{region 'Documentation'}
(*!
<summary>Checks exact finding count and identities; at most one finding per subject.</summary>
*)
{endregion}
METHOD PRIVATE CheckFindings
VAR
    Index : UINT;
    Matches : BOOL;
END_VAR
Index := 1;
FFindingsMatch := TRUE;
Matches := CheckFinding(Subject := FEqual,
    ExpectedResult := FEqualExpectedResult,
    ExpectedFinding := FEqualExpectedFinding,
    Index := Index);
FFindingsMatch := FFindingsMatch AND Matches;
Matches := CheckFinding(Subject := FPattern,
    ExpectedResult := FPatternExpectedResult,
    ExpectedFinding := FPatternExpectedFinding,
    Index := Index);
FFindingsMatch := FFindingsMatch AND Matches;
Matches := CheckFinding(Subject := FAll,
    ExpectedResult := FAllExpectedResult,
    ExpectedFinding := FAllExpectedFinding,
    Index := Index);
FFindingsMatch := FFindingsMatch AND Matches;
Matches := CheckFinding(Subject := FValue,
    ExpectedResult := FValueExpectedResult,
    ExpectedFinding := FValueExpectedFinding,
    Index := Index);
FFindingsMatch := FFindingsMatch AND Matches;
FFindingsMatch := FFindingsMatch
    AND (FCaptureStatus.SequenceId = UINT_TO_UDINT(Index - 1))
    AND (FCaptureStatus.LostEventCount = 0);
END_METHOD

{region 'Documentation'}
(*!
<summary>Rejects incomplete subject, capture or outer Assertion setup.</summary>
*)
{endregion}
METHOD PROTECTED CheckInitialization : BOOL //! TRUE when the inherited initialization check and this concrete fixture check both accept the setup.
CheckInitialization := SUPER^.CheckInitialization();
IF NOT CheckInitialization THEN
    RETURN;
END_IF;

CheckInitialization := FSetupValid
    AND FResults.IsInitialized
    AND FActivity.IsInitialized
    AND FInputs.IsInitialized
    AND FFindings.IsInitialized;
IF NOT CheckInitialization THEN
    EventPublisher.PublishEvent(Event := CreateFrameworkEvent(Name := Name,
        ResourceName := '',
        State := State,
        Severity := E_EventSeverity.Error,
        Message := 'Array selftest setup failed.'));
END_IF;
END_METHOD

{region 'Documentation'}
(*!
<summary>Verifies input preservation without using the tested comparison algorithm.</summary>
*)
{endregion}
METHOD PRIVATE CheckInputs
VAR
    Index : DINT;
    ActualBits : FloatingPointBits_Real;
    SavedBits : FloatingPointBits_Real;
    WideActualBits : FloatingPointBits_LReal;
    WideSavedBits : FloatingPointBits_LReal;
END_VAR
FInputsMatch := TRUE;
FOR Index := -2 TO 1 DO
    ActualBits.Value := FData[Index];
    SavedBits.Value := FDataBefore[Index];
    WideActualBits.Value := FWideData[Index];
    WideSavedBits.Value := FWideDataBefore[Index];
    FInputsMatch := FInputsMatch
        AND (ActualBits.Bits = SavedBits.Bits)
        AND (WideActualBits.Bits = WideSavedBits.Bits);
END_FOR;
FOR Index := 4 TO 5 DO
    ActualBits.Value := FExpected[Index];
    SavedBits.Value := FExpectedBefore[Index];
    FInputsMatch := FInputsMatch AND (ActualBits.Bits = SavedBits.Bits);
END_FOR;
END_METHOD

{region 'Documentation'}
(*!
<summary>Checks literal evaluation results, or NotEvaluated on the reset call.</summary>
*)
{endregion}
METHOD PRIVATE CheckResults
IF FEvaluateSubjects THEN
    FResultsMatch := (FEqual.Result = FEqualExpectedResult)
        AND (FPattern.Result = FPatternExpectedResult)
        AND (FAll.Result = FAllExpectedResult)
        AND (FValue.Result = FValueExpectedResult);
ELSE
    FResultsMatch := (FEqual.Result = E_Result.NotEvaluated)
        AND (FPattern.Result = E_Result.NotEvaluated)
        AND (FAll.Result = E_Result.NotEvaluated)
        AND (FValue.Result = E_Result.NotEvaluated);
END_IF;
FActivityMatch := (FEqual.Enabled = FSubjectEnable)
    AND (FEqual.ObservationActive = (FEvaluateSubjects AND FSubjectEnable))
    AND (FEqual.EvaluationActive = (FEvaluateSubjects AND FSubjectEnable))
    AND (FPattern.Enabled = FSubjectEnable)
    AND (FPattern.ObservationActive = (FEvaluateSubjects AND FSubjectEnable))
    AND (FPattern.EvaluationActive = (FEvaluateSubjects AND FSubjectEnable))
    AND (FAll.Enabled = FSubjectEnable)
    AND (FAll.ObservationActive = (FEvaluateSubjects AND FSubjectEnable))
    AND (FAll.EvaluationActive = (FEvaluateSubjects AND FSubjectEnable))
    AND (FValue.Enabled = FSubjectEnable)
    AND (FValue.ObservationActive = (FEvaluateSubjects AND FSubjectEnable))
    AND (FValue.EvaluationActive = (FEvaluateSubjects AND FSubjectEnable));
END_METHOD

{region 'Documentation'}
(*!
<summary>Initializes outer checks and isolates intentional subject findings.</summary>
*)
{endregion}
METHOD PROTECTED Configure
VAR
    Initialized : BOOL;
END_VAR
FPreparationStateCount := 0;
FTestStateCount := 1;
FResults.Initialize(Parent := THIS^,
    AssertionName := 'Results');
FActivity.Initialize(Parent := THIS^,
    AssertionName := 'Activity');
FInputs.Initialize(Parent := THIS^,
    AssertionName := 'Inputs');
FFindings.Initialize(Parent := THIS^,
    AssertionName := 'Findings');
FSetupValid := FCapture.Initialize(Buffer := FEvents,
    FifoControl := FCaptureFifo,
    Status := FCaptureStatus);
FEqual.BindPublisher(Publisher := FCapture);
Initialized := FEqual.Initialize(Parent := THIS^,
    AssertionName := 'Equal');
FSetupValid := FSetupValid AND Initialized;
FPattern.BindPublisher(Publisher := FCapture);
Initialized := FPattern.Initialize(Parent := THIS^,
    AssertionName := 'Pattern');
FSetupValid := FSetupValid AND Initialized;
FAll.BindPublisher(Publisher := FCapture);
Initialized := FAll.Initialize(Parent := THIS^,
    AssertionName := 'All');
FSetupValid := FSetupValid AND Initialized;
FValue.BindPublisher(Publisher := FCapture);
Initialized := FValue.Initialize(Parent := THIS^,
    AssertionName := 'Value');
FSetupValid := FSetupValid AND Initialized;
END_METHOD

{region 'Documentation'}
(*!
<summary>Completes abort; no asynchronous resource is owned.</summary>
*)
{endregion}
METHOD PROTECTED ProcessAbort
VAR_INPUT
    Enable : BOOL; //! Phase permission supplied by the owning Test Case; FALSE does not authorize progression, while observation may continue.
END_VAR
IF Enable THEN
    CompleteAbort();
END_IF;
END_METHOD

{region 'Documentation'}
(*!
<summary>Latches this call's checks before progression is permitted.</summary>
*)
{endregion}
METHOD PROTECTED ProcessAssertions
VAR_INPUT
    Enable : BOOL; //! Phase permission supplied by the owning Test Case; FALSE does not authorize progression, while observation may continue.
END_VAR
VAR
    Check : BOOL;
END_VAR
Check := Enable AND FObservationReady;
FResults(Enable := Check,
    State := State,
    IN := FResultsMatch);
FActivity(Enable := Check,
    State := State,
    IN := FActivityMatch);
FInputs(Enable := Check,
    State := State,
    IN := FInputsMatch);
FFindings(Enable := Check,
    State := State,
    IN := FFindingsMatch);
IF Check THEN
    FChecked := TRUE;
END_IF;
END_METHOD

{region 'Documentation'}
(*!
<summary>No Preparation phase is needed.</summary>
*)
{endregion}
METHOD PROTECTED ProcessPreparations
VAR_INPUT
    // SA0033: Required hook; this test has no Preparation phase.
    {attribute 'analysis' := '-33'}
    Enable : BOOL; //! Phase permission supplied by the owning Test Case; FALSE does not authorize progression, while observation may continue.
END_VAR
END_METHOD

{region 'Documentation'}
(*!
<summary>Restarts the scenario sequence and outer checks.</summary>
*)
{endregion}
METHOD PROTECTED ProcessReset
FScenario := ScenarioFiniteEqual;
FChecked := FALSE;
FSubjectEnable := FALSE;
FEvaluateSubjects := FALSE;
FObservationReady := FALSE;
FFirstFailedScenario := 0;
FFailedDuringEvaluation := FALSE;
FCapture.Reset();
ResetSubjects();
FResults.Reset();
FActivity.Reset();
FInputs.Reset();
FFindings.Reset();
CompleteReset();
END_METHOD

{region 'Documentation'}
(*!
<summary>Consumes reset, evaluates, then waits for the outer checks before advancing.</summary>
*)
{endregion}
METHOD PROTECTED ProcessTests
VAR_INPUT
    Enable : BOOL; //! Phase permission supplied by the owning Test Case; FALSE does not authorize progression, while observation may continue.
END_VAR
IF NOT Enable THEN
    RETURN;
END_IF;

IF FChecked THEN
    FChecked := FALSE;
    FObservationReady := FALSE;
    IF FEvaluateSubjects THEN
        IF FScenario = LastScenario THEN
            CompleteTests();
            RETURN;
        END_IF;
        FScenario := FScenario + 1;
    END_IF;
    FEvaluateSubjects := NOT FEvaluateSubjects;
END_IF;

IF NOT SelectScenario() THEN
    RETURN;
END_IF;
FCapture.Reset();
IF NOT FEvaluateSubjects THEN
    ResetSubjects();
END_IF;
FDataBefore := FData;
FExpectedBefore := FExpected;
FWideDataBefore := FWideData;

CallSubjects();
CheckResults();
CheckInputs();
CheckFindings();
IF (FFirstFailedScenario = 0)
    AND NOT (FResultsMatch AND FActivityMatch AND FInputsMatch AND FFindingsMatch) THEN
    FFirstFailedScenario := FScenario;
    FFailedDuringEvaluation := FEvaluateSubjects;
END_IF;
FObservationReady := TRUE;
END_METHOD

{region 'Documentation'}
(*!
<summary>Queues reset; the next bound FB call consumes it without evaluating.</summary>
*)
{endregion}
METHOD PRIVATE ResetSubjects
FEqual.Reset();
FPattern.Reset();
FAll.Reset();
FValue.Reset();
END_METHOD

{region 'Documentation'}
(*!
<summary>Selects explicit stimuli and expected results for one scenario.</summary>
*)
{endregion}
METHOD PRIVATE SelectScenario : BOOL //! TRUE after selecting a supported scenario and its literal expectations; FALSE reports an unknown scenario.
VAR
    Index : DINT;
END_VAR
SelectScenario := FALSE;
FSubjectEnable := TRUE;
FQuietNaN.Bits := QuietNaNBits;
FPositiveInfinity.Bits := PositiveInfinityBits;
FNegativeInfinity.Bits := NegativeInfinityBits;
FWideQuietNaN.Bits := WideQuietNaNBits;
FWidePositiveInfinity.Bits := WidePositiveInfinityBits;
FWideNegativeInfinity.Bits := WideNegativeInfinityBits;
FActual := 1.0;
FReference := 1.0;
FWideActual := 1.0;
FWideExpected := 1.0;
FTolerance := 0.0;
FWideTolerance := 0.0;
CASE FScenario OF
    ScenarioFiniteEqual:
        FEqualExpectedResult := E_Result.Passed;
        FEqualExpectedFinding := FALSE;
        FPatternExpectedResult := E_Result.Passed;
        FPatternExpectedFinding := FALSE;
        FAllExpectedResult := E_Result.Passed;
        FAllExpectedFinding := FALSE;
        FValueExpectedResult := E_Result.Passed;
        FValueExpectedFinding := FALSE;
    ScenarioToleranceBoundary:
        FActual := 1.25;
        FWideActual := 1.25;
        FTolerance := 0.25;
        FWideTolerance := 0.25;
        FEqualExpectedResult := E_Result.Passed;
        FEqualExpectedFinding := FALSE;
        FPatternExpectedResult := E_Result.Passed;
        FPatternExpectedFinding := FALSE;
        FAllExpectedResult := E_Result.Passed;
        FAllExpectedFinding := FALSE;
        FValueExpectedResult := E_Result.Passed;
        FValueExpectedFinding := FALSE;
    ScenarioOutsideTolerance:
        FActual := 1.5;
        FWideActual := 1.5;
        FTolerance := 0.25;
        FWideTolerance := 0.25;
        FEqualExpectedResult := E_Result.Failed;
        FEqualExpectedFinding := TRUE;
        FPatternExpectedResult := E_Result.Failed;
        FPatternExpectedFinding := TRUE;
        FAllExpectedResult := E_Result.Failed;
        FAllExpectedFinding := TRUE;
        FValueExpectedResult := E_Result.Failed;
        FValueExpectedFinding := TRUE;
    ScenarioNaNBeforeValidMatch:
        FEqualExpectedResult := E_Result.Failed;
        FEqualExpectedFinding := TRUE;
        FPatternExpectedResult := E_Result.Passed;
        FPatternExpectedFinding := FALSE;
        FAllExpectedResult := E_Result.Failed;
        FAllExpectedFinding := TRUE;
        FValueExpectedResult := E_Result.Passed;
        FValueExpectedFinding := FALSE;
    ScenarioOnlyNaNActual:
        FActual := FQuietNaN.Value;
        FWideActual := FWideQuietNaN.Value;
        FEqualExpectedResult := E_Result.Failed;
        FEqualExpectedFinding := TRUE;
        FPatternExpectedResult := E_Result.Failed;
        FPatternExpectedFinding := TRUE;
        FAllExpectedResult := E_Result.Failed;
        FAllExpectedFinding := TRUE;
        FValueExpectedResult := E_Result.Failed;
        FValueExpectedFinding := TRUE;
    ScenarioPositiveInfinityMatch:
        FActual := FPositiveInfinity.Value;
        FReference := FPositiveInfinity.Value;
        FWideActual := FWidePositiveInfinity.Value;
        FWideExpected := FWidePositiveInfinity.Value;
        FEqualExpectedResult := E_Result.Error;
        FEqualExpectedFinding := TRUE;
        FPatternExpectedResult := E_Result.Passed;
        FPatternExpectedFinding := FALSE;
        FAllExpectedResult := E_Result.Passed;
        FAllExpectedFinding := FALSE;
        FValueExpectedResult := E_Result.Passed;
        FValueExpectedFinding := FALSE;
    ScenarioNegativeInfinityMatch:
        FActual := FNegativeInfinity.Value;
        FReference := FNegativeInfinity.Value;
        FWideActual := FWideNegativeInfinity.Value;
        FWideExpected := FWideNegativeInfinity.Value;
        FEqualExpectedResult := E_Result.Error;
        FEqualExpectedFinding := TRUE;
        FPatternExpectedResult := E_Result.Passed;
        FPatternExpectedFinding := FALSE;
        FAllExpectedResult := E_Result.Passed;
        FAllExpectedFinding := FALSE;
        FValueExpectedResult := E_Result.Passed;
        FValueExpectedFinding := FALSE;
    ScenarioOppositeInfinities:
        FActual := FPositiveInfinity.Value;
        FReference := FNegativeInfinity.Value;
        FWideActual := FWidePositiveInfinity.Value;
        FWideExpected := FWideNegativeInfinity.Value;
        FEqualExpectedResult := E_Result.Error;
        FEqualExpectedFinding := TRUE;
        FPatternExpectedResult := E_Result.Failed;
        FPatternExpectedFinding := TRUE;
        FAllExpectedResult := E_Result.Failed;
        FAllExpectedFinding := TRUE;
        FValueExpectedResult := E_Result.Failed;
        FValueExpectedFinding := TRUE;
    ScenarioPositiveInfinityActual:
        FActual := FPositiveInfinity.Value;
        FWideActual := FWidePositiveInfinity.Value;
        FEqualExpectedResult := E_Result.Failed;
        FEqualExpectedFinding := TRUE;
        FPatternExpectedResult := E_Result.Failed;
        FPatternExpectedFinding := TRUE;
        FAllExpectedResult := E_Result.Failed;
        FAllExpectedFinding := TRUE;
        FValueExpectedResult := E_Result.Failed;
        FValueExpectedFinding := TRUE;
    ScenarioNegativeInfinityActual:
        FActual := FNegativeInfinity.Value;
        FWideActual := FWideNegativeInfinity.Value;
        FEqualExpectedResult := E_Result.Failed;
        FEqualExpectedFinding := TRUE;
        FPatternExpectedResult := E_Result.Failed;
        FPatternExpectedFinding := TRUE;
        FAllExpectedResult := E_Result.Failed;
        FAllExpectedFinding := TRUE;
        FValueExpectedResult := E_Result.Failed;
        FValueExpectedFinding := TRUE;
    ScenarioNaNExpected:
        FReference := FQuietNaN.Value;
        FWideExpected := FWideQuietNaN.Value;
        FEqualExpectedResult := E_Result.Error;
        FEqualExpectedFinding := TRUE;
        FPatternExpectedResult := E_Result.Error;
        FPatternExpectedFinding := TRUE;
        FAllExpectedResult := E_Result.Error;
        FAllExpectedFinding := TRUE;
        FValueExpectedResult := E_Result.Error;
        FValueExpectedFinding := TRUE;
    ScenarioLateNaNExpected:
        FEqualExpectedResult := E_Result.Error;
        FEqualExpectedFinding := TRUE;
        FPatternExpectedResult := E_Result.Error;
        FPatternExpectedFinding := TRUE;
        FAllExpectedResult := E_Result.Passed;
        FAllExpectedFinding := FALSE;
        FValueExpectedResult := E_Result.Passed;
        FValueExpectedFinding := FALSE;
    ScenarioNegativeTolerance:
        FTolerance := -0.25;
        FWideTolerance := -0.25;
        FEqualExpectedResult := E_Result.Error;
        FEqualExpectedFinding := TRUE;
        FPatternExpectedResult := E_Result.Error;
        FPatternExpectedFinding := TRUE;
        FAllExpectedResult := E_Result.Error;
        FAllExpectedFinding := TRUE;
        FValueExpectedResult := E_Result.Error;
        FValueExpectedFinding := TRUE;
    ScenarioNaNTolerance:
        FTolerance := FQuietNaN.Value;
        FWideTolerance := FWideQuietNaN.Value;
        FEqualExpectedResult := E_Result.Error;
        FEqualExpectedFinding := TRUE;
        FPatternExpectedResult := E_Result.Error;
        FPatternExpectedFinding := TRUE;
        FAllExpectedResult := E_Result.Error;
        FAllExpectedFinding := TRUE;
        FValueExpectedResult := E_Result.Error;
        FValueExpectedFinding := TRUE;
    ScenarioInfiniteTolerance:
        FTolerance := FPositiveInfinity.Value;
        FWideTolerance := FWidePositiveInfinity.Value;
        FEqualExpectedResult := E_Result.Error;
        FEqualExpectedFinding := TRUE;
        FPatternExpectedResult := E_Result.Error;
        FPatternExpectedFinding := TRUE;
        FAllExpectedResult := E_Result.Error;
        FAllExpectedFinding := TRUE;
        FValueExpectedResult := E_Result.Error;
        FValueExpectedFinding := TRUE;
ELSE
    Error(Message := 'Unknown array Assertion scenario.');
    RETURN;
END_CASE;
FOR Index := -2 TO 1 DO
    FData[Index] := FActual;
    FWideData[Index] := FWideActual;
END_FOR;
FExpected[4] := FReference;
FExpected[5] := FReference;
IF FScenario = ScenarioNaNBeforeValidMatch THEN
    FData[-2] := FQuietNaN.Value;
    FWideData[-2] := FWideQuietNaN.Value;
END_IF;
IF FScenario = ScenarioLateNaNExpected THEN
    FExpected[5] := FQuietNaN.Value;
    FData[-2] := 9.0;
END_IF;
SelectScenario := TRUE;
END_METHOD

END_FUNCTION_BLOCK

// ---- Framework/Assertions/POU/Arrays/Real/AssertEqualArray_Real.TcPOU
{region 'Documentation'}
(*!
<summary>Compares the entire Expected array with IN starting at StartIndex.</summary>
<description>

StartIndex is an absolute declared IN index. The entire Expected array, starting at its
own lower bound, determines the compared length and must fit IN. Invalid references or ranges
report Error.

Keep supplied arrays stable for the call. Input data is read, not copied or retained as a
snapshot.

Every Expected element must be finite; otherwise Error. A non-finite actual element is a
mismatch (Failed), not an invalid Expected value.

Tolerance is absolute, in the same units as the values, finite and non-negative. Its
default zero requests exact comparison. The equality boundary is inclusive; larger differences
are unequal. Difference checking avoids overflow for large finite operands.

Numeric diagnostics use the formatter's default six significant digits; rounding affects
the message only, not the comparison.

</description>
*)
{endregion}
FUNCTION_BLOCK AssertEqualArray_Real EXTENDS AssertionBase
VAR_INPUT
    Tolerance : REAL := 0.0; //! Maximum absolute allowed difference; finite and non-negative.
    StartIndex : DINT; //! First compared index in IN; Expected starts at its own lower bound.
END_VAR
VAR_IN_OUT CONSTANT
    IN : ARRAY[*] OF REAL; //! Read-only actual data; the selected range must remain stable during the call.
    Expected : ARRAY[*] OF REAL; //! Read-only expected sequence starting at its own lower bound; must fit the selected actual range.
END_VAR

SUPER^();

{region 'Documentation'}
(*!
<summary>Validate the selected range and expectations before comparing elements.</summary>
*)
{endregion}
METHOD PROTECTED Assert
VAR
    ReferenceValue : REAL;
    ValuesEqual : BOOL;
    Value : REAL;
    InLowerIndex : DINT;
    InUpperIndex : DINT;
    ExpectedLowerIndex : DINT;
    ExpectedUpperIndex : DINT;
    ExpectedLength : LINT;
    EndIndex : LINT;
    Offset : LINT;
    InIndex : DINT;
    ExpectedIndex : DINT;
    Message : STRING(GVL_Constants.MessageLength);
    ExpectedText : STRING(GVL_Constants.AssertionValueLength);
    ActualText : STRING(GVL_Constants.AssertionValueLength);
END_VAR
IF NOT EvaluationActive THEN
    RETURN;
END_IF;

IF Result = E_Result.Error THEN
    RETURN;
END_IF;

// C0371: FB inputs are checked here before any reference access.
{warning disable C0371}
IF NOT __ISVALIDREF(IN) THEN
    Error(Message := 'Assertion error: IN reference is invalid.');
    RETURN;
END_IF;

IF NOT __ISVALIDREF(Expected) THEN
    Error(Message := 'Assertion error: Expected reference is invalid.');
    RETURN;
END_IF;

IF NOT Tc2_Utilities.RealIsFinite(x := Tolerance) THEN
    Error(Message := 'Assertion error: Tolerance must be finite.');
    RETURN;
END_IF;

IF Tolerance < 0.0 THEN
    Error(Message := 'Assertion error: Tolerance must not be negative.');
    RETURN;
END_IF;

InLowerIndex := LOWER_BOUND(IN, 1);
InUpperIndex := UPPER_BOUND(IN, 1);
ExpectedLowerIndex := LOWER_BOUND(Expected, 1);
ExpectedUpperIndex := UPPER_BOUND(Expected, 1);
ExpectedLength := DINT_TO_LINT(ExpectedUpperIndex) - DINT_TO_LINT(ExpectedLowerIndex) + 1;
EndIndex := DINT_TO_LINT(StartIndex) + ExpectedLength - 1;

IF (ExpectedLength <= 0)
    OR (StartIndex < InLowerIndex) OR (StartIndex > InUpperIndex)
    OR (EndIndex > DINT_TO_LINT(InUpperIndex)) THEN
    Message := CONCAT('Assertion error: array range is invalid. StartIndex = ',
        DINT_TO_STRING(StartIndex));
    Message := CONCAT(Message, ', EndIndex = ');
    Message := CONCAT(Message, LINT_TO_STRING(EndIndex));
    Message := CONCAT(Message, ', InLowerIndex = ');
    Message := CONCAT(Message, DINT_TO_STRING(InLowerIndex));
    Message := CONCAT(Message, ', InUpperIndex = ');
    Message := CONCAT(Message, DINT_TO_STRING(InUpperIndex));
    Message := CONCAT(Message, ', ExpectedLength = ');
    Message := CONCAT(Message, LINT_TO_STRING(ExpectedLength));
    Message := CONCAT(Message, '.');
    Error(Message := Message);
    RETURN;
END_IF;

FOR Offset := 0 TO ExpectedLength - 1 DO
    ExpectedIndex := LINT_TO_DINT(DINT_TO_LINT(ExpectedLowerIndex) + Offset);
    Value := Expected[ExpectedIndex];
    IF NOT Tc2_Utilities.RealIsFinite(x := Value) THEN
        Message := CONCAT('Assertion error: Expected element must be finite. Index = ',
            DINT_TO_STRING(ExpectedIndex));
        Message := CONCAT(Message, '.');
        Error(Message := Message);
        RETURN;
    END_IF;
END_FOR;

IF Result = E_Result.Failed THEN
    RETURN;
END_IF;

FOR Offset := 0 TO ExpectedLength - 1 DO
    InIndex := LINT_TO_DINT(DINT_TO_LINT(StartIndex) + Offset);
    ExpectedIndex := LINT_TO_DINT(DINT_TO_LINT(ExpectedLowerIndex) + Offset);
    Value := IN[InIndex];
    ReferenceValue := Expected[ExpectedIndex];
    ValuesEqual := FALSE;
    IF NOT Tc2_Utilities.RealIsNaN(x := Value) THEN
        IF Value = ReferenceValue THEN
            ValuesEqual := TRUE;
        ELSIF Tc2_Utilities.RealIsFinite(x := Value)
            AND Tc2_Utilities.RealIsFinite(x := ReferenceValue) THEN
            ValuesEqual := IsWithinTolerance_Real(IN := Value,
                Expected := ReferenceValue,
                Tolerance := Tolerance);
        END_IF;
    END_IF;
    IF NOT ValuesEqual THEN
        ExpectedText := CreateAssertionTextValue_Real(Value := Expected[ExpectedIndex]);
        Value := IN[InIndex];
        IF Tc2_Utilities.RealIsFinite(x := Value) THEN
            ActualText := CreateAssertionTextValue_Real(Value := IN[InIndex]);
        ELSE
            ActualText := '<non-finite>';
        END_IF;
        Message := CONCAT('Assertion failed: array elements differ. Expected[',
            DINT_TO_STRING(ExpectedIndex));
        Message := CONCAT(Message, '] = ');
        Message := CONCAT(Message, ExpectedText);
        Message := CONCAT(Message, ', IN[');
        Message := CONCAT(Message, DINT_TO_STRING(InIndex));
        Message := CONCAT(Message, '] = ');
        Message := CONCAT(Message, ActualText);
        Message := CONCAT(Message, '.');
        Message := CONCAT(Message, ' Tolerance = ');
        Message := CONCAT(Message, CreateAssertionTextValue_Real(Value := Tolerance));
        Fail(Message := Message);
        RETURN;
    END_IF;
END_FOR;

Pass();
{warning restore C0371}
END_METHOD

END_FUNCTION_BLOCK

// ---- Framework/Assertions/POU/Arrays/Real/AssertArrayContainsArray_Real.TcPOU
{region 'Documentation'}
(*!
<summary>Searches the selected IN range for the complete contiguous Expected pattern.</summary>
<description>

StartIndex is an absolute declared IN index, not an offset. Length selects 1..255
elements; the complete selected range must fit IN. Invalid references or ranges report
Error.

Keep supplied arrays stable for the call. Input data is read, not copied or retained as a
snapshot.

The complete Expected pattern must be nonempty and fit the selected IN range; an
oversized pattern reports Error, not a missing-match result.

Expected must not contain NaN (Error), but may contain either infinity. Actual NaN never
matches; equal signed infinities match. Non-finite data elsewhere in a search does not
invalidate the entire range.

Tolerance is absolute, in the same units as the values, finite and non-negative. Its
default zero requests exact comparison. The equality boundary is inclusive; larger differences
are unequal. Difference checking avoids overflow for large finite operands.

Numeric diagnostics use the formatter's default six significant digits; rounding affects
the message only, not the comparison.

</description>
*)
{endregion}
FUNCTION_BLOCK AssertArrayContainsArray_Real EXTENDS AssertionBase
VAR_INPUT
    StartIndex : DINT; //! First selected index in IN; uses the array's declared index range, not a zero-based offset.
    Length : USINT; //! Number of searched elements, from 1 through 255.
    Tolerance : REAL := 0.0; //! Maximum absolute difference accepted as equal; must be finite and non-negative.
END_VAR
VAR_IN_OUT CONSTANT
    IN : ARRAY[*] OF REAL; //! Read-only search data; keep stable during the call.
    Expected : ARRAY[*] OF REAL; //! Read-only expected sequence starting at its own lower bound; must fit the selected actual range.
END_VAR

SUPER^();

{region 'Documentation'}
(*!
<summary>Validate configuration before searching the selected range.</summary>
*)
{endregion}
METHOD PROTECTED Assert
VAR
    InLowerIndex : DINT;
    InUpperIndex : DINT;
    EndIndex : LINT;
    Offset : LINT;
    InIndex : DINT;
    ExpectedLowerIndex : DINT;
    ExpectedUpperIndex : DINT;
    ExpectedLength : LINT;
    ExpectedIndex : DINT;
    CandidateOffset : LINT;
    PatternFound : BOOL;
    PatternMatches : BOOL;
    ValuesEqual : BOOL;
    ExpectedValue : REAL;
    Message : STRING(GVL_Constants.MessageLength);
    Value : REAL;
END_VAR
IF NOT EvaluationActive THEN
    RETURN;
END_IF;

IF Result = E_Result.Error THEN
    RETURN;
END_IF;

// C0371: FB input is checked here before any reference access.
{warning disable C0371}
IF NOT __ISVALIDREF(IN) THEN
    Error(Message := 'Assertion error: IN reference is invalid.');
    RETURN;
END_IF;

IF NOT Tc2_Utilities.RealIsFinite(x := Tolerance) THEN
    Error(Message := 'Assertion error: Tolerance must be finite.');
    RETURN;
END_IF;

IF Tolerance < 0.0 THEN
    Error(Message := 'Assertion error: Tolerance must not be negative.');
    RETURN;
END_IF;

IF NOT __ISVALIDREF(Expected) THEN
    Error(Message := 'Assertion error: Expected reference is invalid.');
    RETURN;
END_IF;

InLowerIndex := LOWER_BOUND(IN, 1);
InUpperIndex := UPPER_BOUND(IN, 1);
EndIndex := DINT_TO_LINT(StartIndex) + USINT_TO_LINT(Length) - 1;

ExpectedLowerIndex := LOWER_BOUND(Expected, 1);
ExpectedUpperIndex := UPPER_BOUND(Expected, 1);
ExpectedLength := DINT_TO_LINT(ExpectedUpperIndex) - DINT_TO_LINT(ExpectedLowerIndex) + 1;

IF (Length = 0)
    OR (ExpectedLength <= 0) OR (ExpectedLength > USINT_TO_LINT(Length))
    OR (StartIndex < InLowerIndex) OR (StartIndex > InUpperIndex)
    OR (EndIndex > DINT_TO_LINT(InUpperIndex)) THEN
    Message := CONCAT('Assertion error: array range or pattern is invalid. StartIndex = ',
        DINT_TO_STRING(StartIndex));
    Message := CONCAT(Message, ', Length = ');
    Message := CONCAT(Message, USINT_TO_STRING(Length));
    Message := CONCAT(Message, ', ExpectedLength = ');
    Message := CONCAT(Message, LINT_TO_STRING(ExpectedLength));
    Message := CONCAT(Message, '.');
    Error(Message := Message);
    RETURN;
END_IF;

FOR Offset := 0 TO ExpectedLength - 1 DO
    ExpectedIndex := LINT_TO_DINT(DINT_TO_LINT(ExpectedLowerIndex) + Offset);
    ExpectedValue := Expected[ExpectedIndex];
    IF Tc2_Utilities.RealIsNaN(x := ExpectedValue) THEN
        Message := CONCAT('Assertion error: Expected must not contain NaN. Index = ',
            DINT_TO_STRING(ExpectedIndex));
        Error(Message := Message);
        RETURN;
    END_IF;
END_FOR;

IF Result = E_Result.Failed THEN
    RETURN;
END_IF;

PatternFound := FALSE;
FOR CandidateOffset := 0 TO USINT_TO_LINT(Length) - ExpectedLength DO
    PatternMatches := TRUE;
    FOR Offset := 0 TO ExpectedLength - 1 DO
        InIndex := LINT_TO_DINT(DINT_TO_LINT(StartIndex) + CandidateOffset + Offset);
        ExpectedIndex := LINT_TO_DINT(DINT_TO_LINT(ExpectedLowerIndex) + Offset);
        Value := IN[InIndex];
        ExpectedValue := Expected[ExpectedIndex];
        ValuesEqual := FALSE;
        IF NOT Tc2_Utilities.RealIsNaN(x := Value) THEN
            IF Value = ExpectedValue THEN
                ValuesEqual := TRUE;
            ELSIF Tc2_Utilities.RealIsFinite(x := Value)
                AND Tc2_Utilities.RealIsFinite(x := ExpectedValue) THEN
                ValuesEqual := IsWithinTolerance_Real(IN := Value,
                    Expected := ExpectedValue,
                    Tolerance := Tolerance);
            END_IF;
        END_IF;
        IF NOT ValuesEqual THEN
            PatternMatches := FALSE;
            EXIT;
        END_IF;
    END_FOR;

    IF PatternMatches THEN
        PatternFound := TRUE;
        EXIT;
    END_IF;
END_FOR;

IF NOT PatternFound THEN
    Message := CONCAT('Assertion failed: array range does not contain Expected pattern. ExpectedRange = [',
        DINT_TO_STRING(ExpectedLowerIndex));
    Message := CONCAT(Message, '..');
    Message := CONCAT(Message, DINT_TO_STRING(ExpectedUpperIndex));
    Message := CONCAT(Message, '], ActualRange = [');
    Message := CONCAT(Message, DINT_TO_STRING(StartIndex));
    Message := CONCAT(Message, '..');
    Message := CONCAT(Message, LINT_TO_STRING(EndIndex));
    Message := CONCAT(Message, ']');
    Message := CONCAT(Message, ', Tolerance = ');
    Message := CONCAT(Message, CreateAssertionTextValue_Real(Value := Tolerance));
    Message := CONCAT(Message, '.');
    Fail(Message := Message);
    RETURN;
END_IF;

Pass();
{warning restore C0371}
END_METHOD

END_FUNCTION_BLOCK

// ---- Framework/Assertions/POU/Arrays/LReal/AssertArrayAllEqual_LReal.TcPOU
{region 'Documentation'}
(*!
<summary>Checks every selected IN element against Expected; reports the first
mismatch.</summary>
<description>

StartIndex is an absolute declared IN index, not an offset. Length selects 1..255
elements; the complete selected range must fit IN. Invalid references or ranges report
Error.

Keep supplied arrays stable for the call. Input data is read, not copied or retained as a
snapshot.

Expected must not contain NaN (Error), but may contain either infinity. Actual NaN never
matches; equal signed infinities match. Non-finite data elsewhere in a search does not
invalidate the entire range.

Tolerance is absolute, in the same units as the values, finite and non-negative. Its
default zero requests exact comparison. The equality boundary is inclusive; larger differences
are unequal. Difference checking avoids overflow for large finite operands.

Numeric diagnostics use the formatter's default six significant digits; rounding affects
the message only, not the comparison.

</description>
*)
{endregion}
FUNCTION_BLOCK AssertArrayAllEqual_LReal EXTENDS AssertionBase
VAR_INPUT
    StartIndex : DINT; //! First selected index in IN; uses the array's declared index range, not a zero-based offset.
    Length : USINT; //! Number of compared elements, from 1 through 255.
    Expected : LREAL; //! Reference value for comparison with IN.
    Tolerance : LREAL := 0.0; //! Maximum absolute difference accepted as equal; must be finite and non-negative.
END_VAR
VAR_IN_OUT CONSTANT
    IN : ARRAY[*] OF LREAL; //! Read-only compared data; keep stable during the call.
END_VAR

SUPER^();

{region 'Documentation'}
(*!
<summary>Validate configuration before comparing the selected range.</summary>
*)
{endregion}
METHOD PROTECTED Assert
VAR
    InLowerIndex : DINT;
    InUpperIndex : DINT;
    EndIndex : LINT;
    Offset : LINT;
    InIndex : DINT;
    ValuesEqual : BOOL;
    Message : STRING(GVL_Constants.MessageLength);
    ActualText : STRING(GVL_Constants.AssertionValueLength);
    ExpectedText : STRING(GVL_Constants.AssertionValueLength);
    Value : LREAL;
END_VAR
IF NOT EvaluationActive THEN
    RETURN;
END_IF;

IF Result = E_Result.Error THEN
    RETURN;
END_IF;

// C0371: FB input is checked here before any reference access.
{warning disable C0371}
IF NOT __ISVALIDREF(IN) THEN
    Error(Message := 'Assertion error: IN reference is invalid.');
    RETURN;
END_IF;

IF Tc2_Utilities.LrealIsNaN(x := Expected) THEN
    Error(Message := 'Assertion error: Expected must not be NaN.');
    RETURN;
END_IF;

IF NOT Tc2_Utilities.LrealIsFinite(x := Tolerance) THEN
    Error(Message := 'Assertion error: Tolerance must be finite.');
    RETURN;
END_IF;

IF Tolerance < 0.0 THEN
    Error(Message := 'Assertion error: Tolerance must not be negative.');
    RETURN;
END_IF;

InLowerIndex := LOWER_BOUND(IN, 1);
InUpperIndex := UPPER_BOUND(IN, 1);
EndIndex := DINT_TO_LINT(StartIndex) + USINT_TO_LINT(Length) - 1;

IF (Length = 0)
    OR (StartIndex < InLowerIndex) OR (StartIndex > InUpperIndex)
    OR (EndIndex > DINT_TO_LINT(InUpperIndex)) THEN
    Message := CONCAT('Assertion error: array range is invalid. StartIndex = ',
        DINT_TO_STRING(StartIndex));
    Message := CONCAT(Message, ', Length = ');
    Message := CONCAT(Message, USINT_TO_STRING(Length));
    Message := CONCAT(Message, '.');
    Error(Message := Message);
    RETURN;
END_IF;

IF Result = E_Result.Failed THEN
    RETURN;
END_IF;

FOR Offset := 0 TO USINT_TO_LINT(Length) - 1 DO
    InIndex := LINT_TO_DINT(DINT_TO_LINT(StartIndex) + Offset);
    ValuesEqual := FALSE;
    Value := IN[InIndex];
    IF NOT Tc2_Utilities.LrealIsNaN(x := Value) THEN
        IF Value = Expected THEN
            ValuesEqual := TRUE;
        ELSIF Tc2_Utilities.LrealIsFinite(x := Value)
            AND Tc2_Utilities.LrealIsFinite(x := Expected) THEN
            ValuesEqual := IsWithinTolerance_LReal(IN := Value,
                Expected := Expected,
                Tolerance := Tolerance);
        END_IF;
    END_IF;
    IF NOT ValuesEqual THEN
        EXIT;
    END_IF;
END_FOR;

IF NOT ValuesEqual THEN
    IF Tc2_Utilities.LrealIsFinite(x := Expected) THEN
        ExpectedText := CreateAssertionTextValue_LReal(Value := Expected);
    ELSIF Expected > 0.0 THEN
        ExpectedText := '+Infinity';
    ELSE
        ExpectedText := '-Infinity';
    END_IF;
    Value := IN[InIndex];
    IF Tc2_Utilities.LrealIsNaN(x := Value) THEN
        ActualText := 'NaN';
    ELSIF Tc2_Utilities.LrealIsFinite(x := Value) THEN
        ActualText := CreateAssertionTextValue_LReal(Value := Value);
    ELSIF Value > 0.0 THEN
        ActualText := '+Infinity';
    ELSE
        ActualText := '-Infinity';
    END_IF;
    Message := CONCAT('Assertion failed: array value is not equal. Expected = ',
        ExpectedText);
    Message := CONCAT(Message, ', Actual[');
    Message := CONCAT(Message, DINT_TO_STRING(InIndex));
    Message := CONCAT(Message, '] = ');
    Message := CONCAT(Message, ActualText);
    Message := CONCAT(Message, ', Range = [');
    Message := CONCAT(Message, DINT_TO_STRING(StartIndex));
    Message := CONCAT(Message, '..');
    Message := CONCAT(Message, LINT_TO_STRING(EndIndex));
    Message := CONCAT(Message, ']');
    Message := CONCAT(Message, ', Tolerance = ');
    Message := CONCAT(Message, CreateAssertionTextValue_LReal(Value := Tolerance));
    Message := CONCAT(Message, '.');
    Fail(Message := Message);
    RETURN;
END_IF;

Pass();
{warning restore C0371}
END_METHOD

END_FUNCTION_BLOCK

// ---- Framework/Assertions/POU/Arrays/LReal/AssertArrayContainsValue_LReal.TcPOU
{region 'Documentation'}
(*!
<summary>Searches the selected IN range for Expected; invalid configuration reports
Error.</summary>
<description>

StartIndex is an absolute declared IN index, not an offset. Length selects 1..255
elements; the complete selected range must fit IN. Invalid references or ranges report
Error.

Keep supplied arrays stable for the call. Input data is read, not copied or retained as a
snapshot.

Expected must not contain NaN (Error), but may contain either infinity. Actual NaN never
matches; equal signed infinities match. Non-finite data elsewhere in a search does not
invalidate the entire range.

Tolerance is absolute, in the same units as the values, finite and non-negative. Its
default zero requests exact comparison. The equality boundary is inclusive; larger differences
are unequal. Difference checking avoids overflow for large finite operands.

Numeric diagnostics use the formatter's default six significant digits; rounding affects
the message only, not the comparison.

</description>
*)
{endregion}
FUNCTION_BLOCK AssertArrayContainsValue_LReal EXTENDS AssertionBase
VAR_INPUT
    StartIndex : DINT; //! First selected index in IN; uses the array's declared index range, not a zero-based offset.
    Length : USINT; //! Number of searched elements, from 1 through 255.
    Expected : LREAL; //! Reference value for comparison with IN.
    Tolerance : LREAL := 0.0; //! Maximum absolute difference accepted as equal; must be finite and non-negative.
END_VAR
VAR_IN_OUT CONSTANT
    IN : ARRAY[*] OF LREAL; //! Read-only search data; keep stable during the call.
END_VAR

SUPER^();

{region 'Documentation'}
(*!
<summary>Validate configuration before searching the selected range.</summary>
*)
{endregion}
METHOD PROTECTED Assert
VAR
    InLowerIndex : DINT;
    InUpperIndex : DINT;
    EndIndex : LINT;
    Offset : LINT;
    InIndex : DINT;
    ValueFound : BOOL;
    Message : STRING(GVL_Constants.MessageLength);
    ExpectedText : STRING(GVL_Constants.AssertionValueLength);
    Value : LREAL;
END_VAR
IF NOT EvaluationActive THEN
    RETURN;
END_IF;

IF Result = E_Result.Error THEN
    RETURN;
END_IF;

// C0371: FB input is checked here before any reference access.
{warning disable C0371}
IF NOT __ISVALIDREF(IN) THEN
    Error(Message := 'Assertion error: IN reference is invalid.');
    RETURN;
END_IF;

IF Tc2_Utilities.LrealIsNaN(x := Expected) THEN
    Error(Message := 'Assertion error: Expected must not be NaN.');
    RETURN;
END_IF;

IF NOT Tc2_Utilities.LrealIsFinite(x := Tolerance) THEN
    Error(Message := 'Assertion error: Tolerance must be finite.');
    RETURN;
END_IF;

IF Tolerance < 0.0 THEN
    Error(Message := 'Assertion error: Tolerance must not be negative.');
    RETURN;
END_IF;

InLowerIndex := LOWER_BOUND(IN, 1);
InUpperIndex := UPPER_BOUND(IN, 1);
EndIndex := DINT_TO_LINT(StartIndex) + USINT_TO_LINT(Length) - 1;

IF (Length = 0)
    OR (StartIndex < InLowerIndex) OR (StartIndex > InUpperIndex)
    OR (EndIndex > DINT_TO_LINT(InUpperIndex)) THEN
    Message := CONCAT('Assertion error: array range is invalid. StartIndex = ',
        DINT_TO_STRING(StartIndex));
    Message := CONCAT(Message, ', Length = ');
    Message := CONCAT(Message, USINT_TO_STRING(Length));
    Message := CONCAT(Message, '.');
    Error(Message := Message);
    RETURN;
END_IF;

IF Result = E_Result.Failed THEN
    RETURN;
END_IF;

ValueFound := FALSE;
FOR Offset := 0 TO USINT_TO_LINT(Length) - 1 DO
    InIndex := LINT_TO_DINT(DINT_TO_LINT(StartIndex) + Offset);
    Value := IN[InIndex];
    IF NOT Tc2_Utilities.LrealIsNaN(x := Value) THEN
        IF Value = Expected THEN
            ValueFound := TRUE;
        ELSIF Tc2_Utilities.LrealIsFinite(x := Value)
            AND Tc2_Utilities.LrealIsFinite(x := Expected) THEN
            ValueFound := IsWithinTolerance_LReal(IN := Value,
                Expected := Expected,
                Tolerance := Tolerance);
        END_IF;
    END_IF;
    IF ValueFound THEN
        EXIT;
    END_IF;
END_FOR;

IF NOT ValueFound THEN
    IF Tc2_Utilities.LrealIsFinite(x := Expected) THEN
        ExpectedText := CreateAssertionTextValue_LReal(Value := Expected);
    ELSIF Expected > 0.0 THEN
        ExpectedText := '+Infinity';
    ELSE
        ExpectedText := '-Infinity';
    END_IF;
    Message := CONCAT('Assertion failed: array range does not contain Expected = ',
        ExpectedText);
    Message := CONCAT(Message, ', Range = [');
    Message := CONCAT(Message, DINT_TO_STRING(StartIndex));
    Message := CONCAT(Message, '..');
    Message := CONCAT(Message, LINT_TO_STRING(EndIndex));
    Message := CONCAT(Message, ']');
    Message := CONCAT(Message, ', Tolerance = ');
    Message := CONCAT(Message, CreateAssertionTextValue_LReal(Value := Tolerance));
    Message := CONCAT(Message, '.');
    Fail(Message := Message);
    RETURN;
END_IF;

Pass();
{warning restore C0371}
END_METHOD

END_FUNCTION_BLOCK

// ---- SelfTests/TestCases/TestSuite_AssertionArrays/Test_AssertionArrayTextBridge.TcPOU
{region 'Documentation'}
(*!
<summary>Checks BYTE/STRING and WORD/WSTRING comparisons without trimming or stopping at array zero.</summary>
<description>
Each independent scenario consumes a bound reset call before its evaluation call.
ProcessAssertions checks the observation before ProcessTests advances.
SelectScenario holds explicit expected results; no production algorithm is mirrored.
Expected findings remain in the local capture; only outer checks affect the test result.
FirstFailedScenario and FailedDuringEvaluation retain the first mismatch.
The wide text deliberately contains code units above 255 with the same low bytes as ASCII.
Input zero and trailing padding are data, not implicit string termination.
Eight simultaneous subject findings require capture headroom below the AlmostFull threshold.
</description>
*)
{endregion}
FUNCTION_BLOCK Test_AssertionArrayTextBridge EXTENDS TestCaseBase
VAR
    FEqual : AssertArrayEqualString_Byte;
    FEqualExpectedResult : E_Result;
    FEqualExpectedFinding : BOOL;
    FContains : AssertArrayContainsString_Byte;
    FContainsExpectedResult : E_Result;
    FContainsExpectedFinding : BOOL;
    FStartsWith : AssertArrayStartsWithString_Byte;
    FStartsWithExpectedResult : E_Result;
    FStartsWithExpectedFinding : BOOL;
    FEndsWith : AssertArrayEndsWithString_Byte;
    FEndsWithExpectedResult : E_Result;
    FEndsWithExpectedFinding : BOOL;
    FWideEqual : AssertArrayEqualWString_Word;
    FWideEqualExpectedResult : E_Result;
    FWideEqualExpectedFinding : BOOL;
    FWideContains : AssertArrayContainsWString_Word;
    FWideContainsExpectedResult : E_Result;
    FWideContainsExpectedFinding : BOOL;
    FWideStartsWith : AssertArrayStartsWithWString_Word;
    FWideStartsWithExpectedResult : E_Result;
    FWideStartsWithExpectedFinding : BOOL;
    FWideEndsWith : AssertArrayEndsWithWString_Word;
    FWideEndsWithExpectedResult : E_Result;
    FWideEndsWithExpectedFinding : BOOL;
    FData : ARRAY[-2..3] OF BYTE;
    FDataBefore : ARRAY[-2..3] OF BYTE;
    FWideData : ARRAY[-2..3] OF WORD;
    FWideDataBefore : ARRAY[-2..3] OF WORD;
    FExpected : STRING(Param_Assertions.AssertionStringLength);
    FExpectedBefore : STRING(Param_Assertions.AssertionStringLength);
    FWideExpected : WSTRING(Param_Assertions.AssertionWStringLength);
    FWideExpectedBefore : WSTRING(Param_Assertions.AssertionWStringLength);
    FStartIndex : DINT;
    FLength : USINT;
    FSubjectEnable : BOOL;
    FCapture : EventBuffer;
    FEvents : ARRAY[1..CaptureLength] OF ST_Event;
    FCaptureFifo : ST_FifoStatus;
    FCaptureStatus : ST_EventBufferStatus;
    FSetupValid : BOOL;
    FScenario : UINT;
    FChecked : BOOL;
    FEvaluateSubjects : BOOL;
    FObservationReady : BOOL;
    FFirstFailedScenario : UINT;
    FFailedDuringEvaluation : BOOL;
    FResultsMatch : BOOL;
    FResults : AssertTrue;
    FActivityMatch : BOOL;
    FActivity : AssertTrue;
    FInputsMatch : BOOL;
    FInputs : AssertTrue;
    FFindingsMatch : BOOL;
    FFindings : AssertTrue;
END_VAR
VAR CONSTANT
    CaptureLength : UINT := 12;
    ScenarioBothBoundaries : UINT := 1;
    ScenarioExactRegion : UINT := 2;
    ScenarioFirstOnly : UINT := 3;
    ScenarioLastOnly : UINT := 4;
    ScenarioAbsent : UINT := 5;
    ScenarioPartialAtEnd : UINT := 6;
    ScenarioMatchAfterZero : UINT := 7;
    ScenarioTrailingZeroNotPadding : UINT := 8;
    ScenarioTextLongerThanRange : UINT := 9;
    ScenarioEmptyExpected : UINT := 10;
    ScenarioEmptyRange : UINT := 11;
    ScenarioBeyondUpperBound : UINT := 12;
    ScenarioWideHighByteMismatch : UINT := 13;
    ScenarioFailedCandidateThenMatch : UINT := 14;
    LastScenario : UINT := ScenarioFailedCandidateThenMatch;
END_VAR

SUPER^();

{region 'Documentation'}
(*!
<summary>Aggregates only outer checks, not intentionally failing subjects.</summary>
*)
{endregion}
METHOD PROTECTED AggregateResults
VAR_INPUT
    Aggregator : I_ResultAggregator; //! Borrowed result sink owned by the outer Test Case; add this test's checking Assertions without resetting or retaining the sink.
END_VAR
Aggregator.AddProvider(Provider := FResults);
Aggregator.AddProvider(Provider := FActivity);
Aggregator.AddProvider(Provider := FInputs);
Aggregator.AddProvider(Provider := FFindings);
END_METHOD

{region 'Documentation'}
(*!
<summary>Calls each inherited production subject once with caller-owned input storage.</summary>
*)
{endregion}
METHOD PRIVATE CallSubjects
FEqual(Enable := FSubjectEnable,
    State := E_State.Running,
    StartIndex := FStartIndex,
    Length := FLength,
    IN := FData,
    Expected := FExpected);
FContains(Enable := FSubjectEnable,
    State := E_State.Running,
    StartIndex := FStartIndex,
    Length := FLength,
    IN := FData,
    Expected := FExpected);
FStartsWith(Enable := FSubjectEnable,
    State := E_State.Running,
    StartIndex := FStartIndex,
    Length := FLength,
    IN := FData,
    Expected := FExpected);
FEndsWith(Enable := FSubjectEnable,
    State := E_State.Running,
    StartIndex := FStartIndex,
    Length := FLength,
    IN := FData,
    Expected := FExpected);
FWideEqual(Enable := FSubjectEnable,
    State := E_State.Running,
    StartIndex := FStartIndex,
    Length := FLength,
    IN := FWideData,
    Expected := FWideExpected);
FWideContains(Enable := FSubjectEnable,
    State := E_State.Running,
    StartIndex := FStartIndex,
    Length := FLength,
    IN := FWideData,
    Expected := FWideExpected);
FWideStartsWith(Enable := FSubjectEnable,
    State := E_State.Running,
    StartIndex := FStartIndex,
    Length := FLength,
    IN := FWideData,
    Expected := FWideExpected);
FWideEndsWith(Enable := FSubjectEnable,
    State := E_State.Running,
    StartIndex := FStartIndex,
    Length := FLength,
    IN := FWideData,
    Expected := FWideExpected);
END_METHOD

{region 'Documentation'}
(*!
<summary>Checks one subject finding in call order; expected outcomes come from the scenario.</summary>
*)
{endregion}
METHOD PRIVATE CheckFinding : BOOL //! TRUE when the required finding checks pass; calls requiring no finding also succeed.
VAR_INPUT
    Subject : I_Assertion; //! Assertion interface supplying the expected finding identity.
    ExpectedResult : E_Result; //! Independently authored result expected in the captured finding.
    ExpectedFinding : BOOL; //! TRUE when this scenario requires a finding during active evaluation.
END_VAR
VAR_IN_OUT
    Index : UINT; //! One-based next finding index; advanced when this call checks a required finding.
END_VAR
CheckFinding := TRUE;
IF FEvaluateSubjects AND ExpectedFinding THEN
    CheckFinding := (FEvents[Index].SequenceId = UINT_TO_UDINT(Index))
        AND (FEvents[Index].Name = Subject.Name)
        AND (FEvents[Index].OwnerScope = E_OwnerScope.Assertion)
        AND (FEvents[Index].EventType = E_EventType.Result)
        AND (FEvents[Index].State = E_State.Running)
        AND (FEvents[Index].Result = ExpectedResult)
        AND (FEvents[Index].Message <> '');
    Index := Index + 1;
END_IF;
END_METHOD

{region 'Documentation'}
(*!
<summary>Checks exact finding count and identities; at most one finding per subject.</summary>
*)
{endregion}
METHOD PRIVATE CheckFindings
VAR
    Index : UINT;
    Matches : BOOL;
END_VAR
Index := 1;
FFindingsMatch := TRUE;
Matches := CheckFinding(Subject := FEqual,
    ExpectedResult := FEqualExpectedResult,
    ExpectedFinding := FEqualExpectedFinding,
    Index := Index);
FFindingsMatch := FFindingsMatch AND Matches;
Matches := CheckFinding(Subject := FContains,
    ExpectedResult := FContainsExpectedResult,
    ExpectedFinding := FContainsExpectedFinding,
    Index := Index);
FFindingsMatch := FFindingsMatch AND Matches;
Matches := CheckFinding(Subject := FStartsWith,
    ExpectedResult := FStartsWithExpectedResult,
    ExpectedFinding := FStartsWithExpectedFinding,
    Index := Index);
FFindingsMatch := FFindingsMatch AND Matches;
Matches := CheckFinding(Subject := FEndsWith,
    ExpectedResult := FEndsWithExpectedResult,
    ExpectedFinding := FEndsWithExpectedFinding,
    Index := Index);
FFindingsMatch := FFindingsMatch AND Matches;
Matches := CheckFinding(Subject := FWideEqual,
    ExpectedResult := FWideEqualExpectedResult,
    ExpectedFinding := FWideEqualExpectedFinding,
    Index := Index);
FFindingsMatch := FFindingsMatch AND Matches;
Matches := CheckFinding(Subject := FWideContains,
    ExpectedResult := FWideContainsExpectedResult,
    ExpectedFinding := FWideContainsExpectedFinding,
    Index := Index);
FFindingsMatch := FFindingsMatch AND Matches;
Matches := CheckFinding(Subject := FWideStartsWith,
    ExpectedResult := FWideStartsWithExpectedResult,
    ExpectedFinding := FWideStartsWithExpectedFinding,
    Index := Index);
FFindingsMatch := FFindingsMatch AND Matches;
Matches := CheckFinding(Subject := FWideEndsWith,
    ExpectedResult := FWideEndsWithExpectedResult,
    ExpectedFinding := FWideEndsWithExpectedFinding,
    Index := Index);
FFindingsMatch := FFindingsMatch AND Matches;
FFindingsMatch := FFindingsMatch
    AND (FCaptureStatus.SequenceId = UINT_TO_UDINT(Index - 1))
    AND (FCaptureStatus.LostEventCount = 0);
END_METHOD

{region 'Documentation'}
(*!
<summary>Rejects incomplete subject, capture or outer Assertion setup.</summary>
*)
{endregion}
METHOD PROTECTED CheckInitialization : BOOL //! TRUE when the inherited initialization check and this concrete fixture check both accept the setup.
CheckInitialization := SUPER^.CheckInitialization();
IF NOT CheckInitialization THEN
    RETURN;
END_IF;

CheckInitialization := (Param_Assertions.AssertionStringLength >= 2)
    AND (Param_Assertions.AssertionWStringLength >= 2)
    AND FSetupValid
    AND FResults.IsInitialized
    AND FActivity.IsInitialized
    AND FInputs.IsInitialized
    AND FFindings.IsInitialized;
IF NOT CheckInitialization THEN
    EventPublisher.PublishEvent(Event := CreateFrameworkEvent(Name := Name,
        ResourceName := '',
        State := State,
        Severity := E_EventSeverity.Error,
        Message := 'Array selftest setup failed.'));
END_IF;
END_METHOD

{region 'Documentation'}
(*!
<summary>Verifies input preservation without using the tested comparison algorithm.</summary>
*)
{endregion}
METHOD PRIVATE CheckInputs
VAR
    Index : DINT;
END_VAR
FInputsMatch := TRUE;
FOR Index := -2 TO 3 DO
    FInputsMatch := FInputsMatch AND (FData[Index] = FDataBefore[Index]);
END_FOR;
FOR Index := -2 TO 3 DO
    FInputsMatch := FInputsMatch AND (FWideData[Index] = FWideDataBefore[Index]);
END_FOR;
FInputsMatch := FInputsMatch AND (FExpected = FExpectedBefore)
    AND (FWideExpected = FWideExpectedBefore);
END_METHOD

{region 'Documentation'}
(*!
<summary>Checks literal evaluation results, or NotEvaluated on the reset call.</summary>
*)
{endregion}
METHOD PRIVATE CheckResults
IF FEvaluateSubjects THEN
    FResultsMatch := (FEqual.Result = FEqualExpectedResult)
        AND (FContains.Result = FContainsExpectedResult)
        AND (FStartsWith.Result = FStartsWithExpectedResult)
        AND (FEndsWith.Result = FEndsWithExpectedResult)
        AND (FWideEqual.Result = FWideEqualExpectedResult)
        AND (FWideContains.Result = FWideContainsExpectedResult)
        AND (FWideStartsWith.Result = FWideStartsWithExpectedResult)
        AND (FWideEndsWith.Result = FWideEndsWithExpectedResult);
ELSE
    FResultsMatch := (FEqual.Result = E_Result.NotEvaluated)
        AND (FContains.Result = E_Result.NotEvaluated)
        AND (FStartsWith.Result = E_Result.NotEvaluated)
        AND (FEndsWith.Result = E_Result.NotEvaluated)
        AND (FWideEqual.Result = E_Result.NotEvaluated)
        AND (FWideContains.Result = E_Result.NotEvaluated)
        AND (FWideStartsWith.Result = E_Result.NotEvaluated)
        AND (FWideEndsWith.Result = E_Result.NotEvaluated);
END_IF;
FActivityMatch := (FEqual.Enabled = FSubjectEnable)
    AND (FEqual.ObservationActive = (FEvaluateSubjects AND FSubjectEnable))
    AND (FEqual.EvaluationActive = (FEvaluateSubjects AND FSubjectEnable))
    AND (FContains.Enabled = FSubjectEnable)
    AND (FContains.ObservationActive = (FEvaluateSubjects AND FSubjectEnable))
    AND (FContains.EvaluationActive = (FEvaluateSubjects AND FSubjectEnable))
    AND (FStartsWith.Enabled = FSubjectEnable)
    AND (FStartsWith.ObservationActive = (FEvaluateSubjects AND FSubjectEnable))
    AND (FStartsWith.EvaluationActive = (FEvaluateSubjects AND FSubjectEnable))
    AND (FEndsWith.Enabled = FSubjectEnable)
    AND (FEndsWith.ObservationActive = (FEvaluateSubjects AND FSubjectEnable))
    AND (FEndsWith.EvaluationActive = (FEvaluateSubjects AND FSubjectEnable))
    AND (FWideEqual.Enabled = FSubjectEnable)
    AND (FWideEqual.ObservationActive = (FEvaluateSubjects AND FSubjectEnable))
    AND (FWideEqual.EvaluationActive = (FEvaluateSubjects AND FSubjectEnable))
    AND (FWideContains.Enabled = FSubjectEnable)
    AND (FWideContains.ObservationActive = (FEvaluateSubjects AND FSubjectEnable))
    AND (FWideContains.EvaluationActive = (FEvaluateSubjects AND FSubjectEnable))
    AND (FWideStartsWith.Enabled = FSubjectEnable)
    AND (FWideStartsWith.ObservationActive = (FEvaluateSubjects AND FSubjectEnable))
    AND (FWideStartsWith.EvaluationActive = (FEvaluateSubjects AND FSubjectEnable))
    AND (FWideEndsWith.Enabled = FSubjectEnable)
    AND (FWideEndsWith.ObservationActive = (FEvaluateSubjects AND FSubjectEnable))
    AND (FWideEndsWith.EvaluationActive = (FEvaluateSubjects AND FSubjectEnable));
END_METHOD

{region 'Documentation'}
(*!
<summary>Initializes outer checks and isolates intentional subject findings.</summary>
*)
{endregion}
METHOD PROTECTED Configure
VAR
    Initialized : BOOL;
END_VAR
FPreparationStateCount := 0;
FTestStateCount := 1;
FResults.Initialize(Parent := THIS^,
    AssertionName := 'Results');
FActivity.Initialize(Parent := THIS^,
    AssertionName := 'Activity');
FInputs.Initialize(Parent := THIS^,
    AssertionName := 'Inputs');
FFindings.Initialize(Parent := THIS^,
    AssertionName := 'Findings');
FSetupValid := FCapture.Initialize(Buffer := FEvents,
    FifoControl := FCaptureFifo,
    Status := FCaptureStatus);
FEqual.BindPublisher(Publisher := FCapture);
Initialized := FEqual.Initialize(Parent := THIS^,
    AssertionName := 'Equal');
FSetupValid := FSetupValid AND Initialized;
FContains.BindPublisher(Publisher := FCapture);
Initialized := FContains.Initialize(Parent := THIS^,
    AssertionName := 'Contains');
FSetupValid := FSetupValid AND Initialized;
FStartsWith.BindPublisher(Publisher := FCapture);
Initialized := FStartsWith.Initialize(Parent := THIS^,
    AssertionName := 'StartsWith');
FSetupValid := FSetupValid AND Initialized;
FEndsWith.BindPublisher(Publisher := FCapture);
Initialized := FEndsWith.Initialize(Parent := THIS^,
    AssertionName := 'EndsWith');
FSetupValid := FSetupValid AND Initialized;
FWideEqual.BindPublisher(Publisher := FCapture);
Initialized := FWideEqual.Initialize(Parent := THIS^,
    AssertionName := 'WideEqual');
FSetupValid := FSetupValid AND Initialized;
FWideContains.BindPublisher(Publisher := FCapture);
Initialized := FWideContains.Initialize(Parent := THIS^,
    AssertionName := 'WideContains');
FSetupValid := FSetupValid AND Initialized;
FWideStartsWith.BindPublisher(Publisher := FCapture);
Initialized := FWideStartsWith.Initialize(Parent := THIS^,
    AssertionName := 'WideStartsWith');
FSetupValid := FSetupValid AND Initialized;
FWideEndsWith.BindPublisher(Publisher := FCapture);
Initialized := FWideEndsWith.Initialize(Parent := THIS^,
    AssertionName := 'WideEndsWith');
FSetupValid := FSetupValid AND Initialized;
END_METHOD

{region 'Documentation'}
(*!
<summary>Completes abort; no asynchronous resource is owned.</summary>
*)
{endregion}
METHOD PROTECTED ProcessAbort
VAR_INPUT
    Enable : BOOL; //! Phase permission supplied by the owning Test Case; FALSE does not authorize progression, while observation may continue.
END_VAR
IF Enable THEN
    CompleteAbort();
END_IF;
END_METHOD

{region 'Documentation'}
(*!
<summary>Latches this call's checks before progression is permitted.</summary>
*)
{endregion}
METHOD PROTECTED ProcessAssertions
VAR_INPUT
    Enable : BOOL; //! Phase permission supplied by the owning Test Case; FALSE does not authorize progression, while observation may continue.
END_VAR
VAR
    Check : BOOL;
END_VAR
Check := Enable AND FObservationReady;
FResults(Enable := Check,
    State := State,
    IN := FResultsMatch);
FActivity(Enable := Check,
    State := State,
    IN := FActivityMatch);
FInputs(Enable := Check,
    State := State,
    IN := FInputsMatch);
FFindings(Enable := Check,
    State := State,
    IN := FFindingsMatch);
IF Check THEN
    FChecked := TRUE;
END_IF;
END_METHOD

{region 'Documentation'}
(*!
<summary>No Preparation phase is needed.</summary>
*)
{endregion}
METHOD PROTECTED ProcessPreparations
VAR_INPUT
    // SA0033: Required hook; this test has no Preparation phase.
    {attribute 'analysis' := '-33'}
    Enable : BOOL; //! Phase permission supplied by the owning Test Case; FALSE does not authorize progression, while observation may continue.
END_VAR
END_METHOD

{region 'Documentation'}
(*!
<summary>Restarts the scenario sequence and outer checks.</summary>
*)
{endregion}
METHOD PROTECTED ProcessReset
FScenario := ScenarioBothBoundaries;
FChecked := FALSE;
FSubjectEnable := FALSE;
FEvaluateSubjects := FALSE;
FObservationReady := FALSE;
FFirstFailedScenario := 0;
FFailedDuringEvaluation := FALSE;
FCapture.Reset();
ResetSubjects();
FResults.Reset();
FActivity.Reset();
FInputs.Reset();
FFindings.Reset();
CompleteReset();
END_METHOD

{region 'Documentation'}
(*!
<summary>Consumes reset, evaluates, then waits for the outer checks before advancing.</summary>
*)
{endregion}
METHOD PROTECTED ProcessTests
VAR_INPUT
    Enable : BOOL; //! Phase permission supplied by the owning Test Case; FALSE does not authorize progression, while observation may continue.
END_VAR
IF NOT Enable THEN
    RETURN;
END_IF;

IF FChecked THEN
    FChecked := FALSE;
    FObservationReady := FALSE;
    IF FEvaluateSubjects THEN
        IF FScenario = LastScenario THEN
            CompleteTests();
            RETURN;
        END_IF;
        FScenario := FScenario + 1;
    END_IF;
    FEvaluateSubjects := NOT FEvaluateSubjects;
END_IF;

IF NOT SelectScenario() THEN
    RETURN;
END_IF;
FCapture.Reset();
IF NOT FEvaluateSubjects THEN
    ResetSubjects();
END_IF;
FDataBefore := FData;
FWideDataBefore := FWideData;
FExpectedBefore := FExpected;
FWideExpectedBefore := FWideExpected;
CallSubjects();
CheckResults();
CheckInputs();
CheckFindings();
IF (FFirstFailedScenario = 0)
    AND NOT (FResultsMatch AND FActivityMatch AND FInputsMatch AND FFindingsMatch) THEN
    FFirstFailedScenario := FScenario;
    FFailedDuringEvaluation := FEvaluateSubjects;
END_IF;
FObservationReady := TRUE;
END_METHOD

{region 'Documentation'}
(*!
<summary>Queues reset; the next bound FB call consumes it without evaluating.</summary>
*)
{endregion}
METHOD PRIVATE ResetSubjects
FEqual.Reset();
FContains.Reset();
FStartsWith.Reset();
FEndsWith.Reset();
FWideEqual.Reset();
FWideContains.Reset();
FWideStartsWith.Reset();
FWideEndsWith.Reset();
END_METHOD

{region 'Documentation'}
(*!
<summary>Selects explicit stimuli and expected results for one scenario.</summary>
*)
{endregion}
METHOD PRIVATE SelectScenario : BOOL //! TRUE after selecting a supported scenario and its literal expectations; FALSE reports an unknown scenario.
VAR
    Index : DINT;
END_VAR
SelectScenario := FALSE;
FSubjectEnable := TRUE;
FData[-2] := BYTE#16#41;
FData[-1] := BYTE#16#42;
FData[0] := BYTE#16#78;
FData[1] := BYTE#16#78;
FData[2] := BYTE#16#41;
FData[3] := BYTE#16#42;
FWideData[-2] := WORD#16#0141;
FWideData[-1] := WORD#16#0242;
FWideData[0] := WORD#16#0078;
FWideData[1] := WORD#16#0078;
FWideData[2] := WORD#16#0141;
FWideData[3] := WORD#16#0242;
FExpected := 'AB';
FWideExpected := "AB";
FWideExpected[0] := WORD#16#0141;
FWideExpected[1] := WORD#16#0242;
FStartIndex := -2;
FLength := 6;
CASE FScenario OF
    ScenarioBothBoundaries:
        FEqualExpectedResult := E_Result.Failed;
        FEqualExpectedFinding := TRUE;
        FContainsExpectedResult := E_Result.Passed;
        FContainsExpectedFinding := FALSE;
        FStartsWithExpectedResult := E_Result.Passed;
        FStartsWithExpectedFinding := FALSE;
        FEndsWithExpectedResult := E_Result.Passed;
        FEndsWithExpectedFinding := FALSE;
        FWideEqualExpectedResult := E_Result.Failed;
        FWideEqualExpectedFinding := TRUE;
        FWideContainsExpectedResult := E_Result.Passed;
        FWideContainsExpectedFinding := FALSE;
        FWideStartsWithExpectedResult := E_Result.Passed;
        FWideStartsWithExpectedFinding := FALSE;
        FWideEndsWithExpectedResult := E_Result.Passed;
        FWideEndsWithExpectedFinding := FALSE;
    ScenarioExactRegion:
        FLength := 2;
        FEqualExpectedResult := E_Result.Passed;
        FEqualExpectedFinding := FALSE;
        FContainsExpectedResult := E_Result.Passed;
        FContainsExpectedFinding := FALSE;
        FStartsWithExpectedResult := E_Result.Passed;
        FStartsWithExpectedFinding := FALSE;
        FEndsWithExpectedResult := E_Result.Passed;
        FEndsWithExpectedFinding := FALSE;
        FWideEqualExpectedResult := E_Result.Passed;
        FWideEqualExpectedFinding := FALSE;
        FWideContainsExpectedResult := E_Result.Passed;
        FWideContainsExpectedFinding := FALSE;
        FWideStartsWithExpectedResult := E_Result.Passed;
        FWideStartsWithExpectedFinding := FALSE;
        FWideEndsWithExpectedResult := E_Result.Passed;
        FWideEndsWithExpectedFinding := FALSE;
    ScenarioFirstOnly:
        FData[2] := 120;
        FData[3] := 120;
        FWideData[2] := 120;
        FWideData[3] := 120;
        FEqualExpectedResult := E_Result.Failed;
        FEqualExpectedFinding := TRUE;
        FContainsExpectedResult := E_Result.Passed;
        FContainsExpectedFinding := FALSE;
        FStartsWithExpectedResult := E_Result.Passed;
        FStartsWithExpectedFinding := FALSE;
        FEndsWithExpectedResult := E_Result.Failed;
        FEndsWithExpectedFinding := TRUE;
        FWideEqualExpectedResult := E_Result.Failed;
        FWideEqualExpectedFinding := TRUE;
        FWideContainsExpectedResult := E_Result.Passed;
        FWideContainsExpectedFinding := FALSE;
        FWideStartsWithExpectedResult := E_Result.Passed;
        FWideStartsWithExpectedFinding := FALSE;
        FWideEndsWithExpectedResult := E_Result.Failed;
        FWideEndsWithExpectedFinding := TRUE;
    ScenarioLastOnly:
        FData[-2] := 120;
        FData[-1] := 120;
        FWideData[-2] := 120;
        FWideData[-1] := 120;
        FEqualExpectedResult := E_Result.Failed;
        FEqualExpectedFinding := TRUE;
        FContainsExpectedResult := E_Result.Passed;
        FContainsExpectedFinding := FALSE;
        FStartsWithExpectedResult := E_Result.Failed;
        FStartsWithExpectedFinding := TRUE;
        FEndsWithExpectedResult := E_Result.Passed;
        FEndsWithExpectedFinding := FALSE;
        FWideEqualExpectedResult := E_Result.Failed;
        FWideEqualExpectedFinding := TRUE;
        FWideContainsExpectedResult := E_Result.Passed;
        FWideContainsExpectedFinding := FALSE;
        FWideStartsWithExpectedResult := E_Result.Failed;
        FWideStartsWithExpectedFinding := TRUE;
        FWideEndsWithExpectedResult := E_Result.Passed;
        FWideEndsWithExpectedFinding := FALSE;
    ScenarioAbsent:
        FOR Index := -2 TO 3 DO
            FData[Index] := 120;
            FWideData[Index] := 120;
        END_FOR;
        FEqualExpectedResult := E_Result.Failed;
        FEqualExpectedFinding := TRUE;
        FContainsExpectedResult := E_Result.Failed;
        FContainsExpectedFinding := TRUE;
        FStartsWithExpectedResult := E_Result.Failed;
        FStartsWithExpectedFinding := TRUE;
        FEndsWithExpectedResult := E_Result.Failed;
        FEndsWithExpectedFinding := TRUE;
        FWideEqualExpectedResult := E_Result.Failed;
        FWideEqualExpectedFinding := TRUE;
        FWideContainsExpectedResult := E_Result.Failed;
        FWideContainsExpectedFinding := TRUE;
        FWideStartsWithExpectedResult := E_Result.Failed;
        FWideStartsWithExpectedFinding := TRUE;
        FWideEndsWithExpectedResult := E_Result.Failed;
        FWideEndsWithExpectedFinding := TRUE;
    ScenarioPartialAtEnd:
        FOR Index := -2 TO 2 DO
            FData[Index] := 120;
            FWideData[Index] := 120;
        END_FOR;
        FData[3] := BYTE#16#41;
        FWideData[3] := WORD#16#0141;
        FEqualExpectedResult := E_Result.Failed;
        FEqualExpectedFinding := TRUE;
        FContainsExpectedResult := E_Result.Failed;
        FContainsExpectedFinding := TRUE;
        FStartsWithExpectedResult := E_Result.Failed;
        FStartsWithExpectedFinding := TRUE;
        FEndsWithExpectedResult := E_Result.Failed;
        FEndsWithExpectedFinding := TRUE;
        FWideEqualExpectedResult := E_Result.Failed;
        FWideEqualExpectedFinding := TRUE;
        FWideContainsExpectedResult := E_Result.Failed;
        FWideContainsExpectedFinding := TRUE;
        FWideStartsWithExpectedResult := E_Result.Failed;
        FWideStartsWithExpectedFinding := TRUE;
        FWideEndsWithExpectedResult := E_Result.Failed;
        FWideEndsWithExpectedFinding := TRUE;
    ScenarioMatchAfterZero:
        FData[-2] := 0;
        FWideData[-2] := 0;
        FEqualExpectedResult := E_Result.Failed;
        FEqualExpectedFinding := TRUE;
        FContainsExpectedResult := E_Result.Passed;
        FContainsExpectedFinding := FALSE;
        FStartsWithExpectedResult := E_Result.Failed;
        FStartsWithExpectedFinding := TRUE;
        FEndsWithExpectedResult := E_Result.Passed;
        FEndsWithExpectedFinding := FALSE;
        FWideEqualExpectedResult := E_Result.Failed;
        FWideEqualExpectedFinding := TRUE;
        FWideContainsExpectedResult := E_Result.Passed;
        FWideContainsExpectedFinding := FALSE;
        FWideStartsWithExpectedResult := E_Result.Failed;
        FWideStartsWithExpectedFinding := TRUE;
        FWideEndsWithExpectedResult := E_Result.Passed;
        FWideEndsWithExpectedFinding := FALSE;
    ScenarioTrailingZeroNotPadding:
        FLength := 3;
        FData[0] := 0;
        FWideData[0] := 0;
        FEqualExpectedResult := E_Result.Failed;
        FEqualExpectedFinding := TRUE;
        FContainsExpectedResult := E_Result.Passed;
        FContainsExpectedFinding := FALSE;
        FStartsWithExpectedResult := E_Result.Passed;
        FStartsWithExpectedFinding := FALSE;
        FEndsWithExpectedResult := E_Result.Failed;
        FEndsWithExpectedFinding := TRUE;
        FWideEqualExpectedResult := E_Result.Failed;
        FWideEqualExpectedFinding := TRUE;
        FWideContainsExpectedResult := E_Result.Passed;
        FWideContainsExpectedFinding := FALSE;
        FWideStartsWithExpectedResult := E_Result.Passed;
        FWideStartsWithExpectedFinding := FALSE;
        FWideEndsWithExpectedResult := E_Result.Failed;
        FWideEndsWithExpectedFinding := TRUE;
    ScenarioTextLongerThanRange:
        FLength := 1;
        FEqualExpectedResult := E_Result.Failed;
        FEqualExpectedFinding := TRUE;
        FContainsExpectedResult := E_Result.Failed;
        FContainsExpectedFinding := TRUE;
        FStartsWithExpectedResult := E_Result.Failed;
        FStartsWithExpectedFinding := TRUE;
        FEndsWithExpectedResult := E_Result.Failed;
        FEndsWithExpectedFinding := TRUE;
        FWideEqualExpectedResult := E_Result.Failed;
        FWideEqualExpectedFinding := TRUE;
        FWideContainsExpectedResult := E_Result.Failed;
        FWideContainsExpectedFinding := TRUE;
        FWideStartsWithExpectedResult := E_Result.Failed;
        FWideStartsWithExpectedFinding := TRUE;
        FWideEndsWithExpectedResult := E_Result.Failed;
        FWideEndsWithExpectedFinding := TRUE;
    ScenarioEmptyExpected:
        FExpected := '';
        FWideExpected := "";
        FEqualExpectedResult := E_Result.Error;
        FEqualExpectedFinding := TRUE;
        FContainsExpectedResult := E_Result.Error;
        FContainsExpectedFinding := TRUE;
        FStartsWithExpectedResult := E_Result.Error;
        FStartsWithExpectedFinding := TRUE;
        FEndsWithExpectedResult := E_Result.Error;
        FEndsWithExpectedFinding := TRUE;
        FWideEqualExpectedResult := E_Result.Error;
        FWideEqualExpectedFinding := TRUE;
        FWideContainsExpectedResult := E_Result.Error;
        FWideContainsExpectedFinding := TRUE;
        FWideStartsWithExpectedResult := E_Result.Error;
        FWideStartsWithExpectedFinding := TRUE;
        FWideEndsWithExpectedResult := E_Result.Error;
        FWideEndsWithExpectedFinding := TRUE;
    ScenarioEmptyRange:
        FLength := 0;
        FEqualExpectedResult := E_Result.Error;
        FEqualExpectedFinding := TRUE;
        FContainsExpectedResult := E_Result.Error;
        FContainsExpectedFinding := TRUE;
        FStartsWithExpectedResult := E_Result.Error;
        FStartsWithExpectedFinding := TRUE;
        FEndsWithExpectedResult := E_Result.Error;
        FEndsWithExpectedFinding := TRUE;
        FWideEqualExpectedResult := E_Result.Error;
        FWideEqualExpectedFinding := TRUE;
        FWideContainsExpectedResult := E_Result.Error;
        FWideContainsExpectedFinding := TRUE;
        FWideStartsWithExpectedResult := E_Result.Error;
        FWideStartsWithExpectedFinding := TRUE;
        FWideEndsWithExpectedResult := E_Result.Error;
        FWideEndsWithExpectedFinding := TRUE;
    ScenarioBeyondUpperBound:
        FStartIndex := 3;
        FLength := 2;
        FEqualExpectedResult := E_Result.Error;
        FEqualExpectedFinding := TRUE;
        FContainsExpectedResult := E_Result.Error;
        FContainsExpectedFinding := TRUE;
        FStartsWithExpectedResult := E_Result.Error;
        FStartsWithExpectedFinding := TRUE;
        FEndsWithExpectedResult := E_Result.Error;
        FEndsWithExpectedFinding := TRUE;
        FWideEqualExpectedResult := E_Result.Error;
        FWideEqualExpectedFinding := TRUE;
        FWideContainsExpectedResult := E_Result.Error;
        FWideContainsExpectedFinding := TRUE;
        FWideStartsWithExpectedResult := E_Result.Error;
        FWideStartsWithExpectedFinding := TRUE;
        FWideEndsWithExpectedResult := E_Result.Error;
        FWideEndsWithExpectedFinding := TRUE;
    ScenarioWideHighByteMismatch:
        FWideExpected[0] := WORD#16#0241;
        FEqualExpectedResult := E_Result.Failed;
        FEqualExpectedFinding := TRUE;
        FContainsExpectedResult := E_Result.Passed;
        FContainsExpectedFinding := FALSE;
        FStartsWithExpectedResult := E_Result.Passed;
        FStartsWithExpectedFinding := FALSE;
        FEndsWithExpectedResult := E_Result.Passed;
        FEndsWithExpectedFinding := FALSE;
        FWideEqualExpectedResult := E_Result.Failed;
        FWideEqualExpectedFinding := TRUE;
        FWideContainsExpectedResult := E_Result.Failed;
        FWideContainsExpectedFinding := TRUE;
        FWideStartsWithExpectedResult := E_Result.Failed;
        FWideStartsWithExpectedFinding := TRUE;
        FWideEndsWithExpectedResult := E_Result.Failed;
        FWideEndsWithExpectedFinding := TRUE;
    ScenarioFailedCandidateThenMatch:
        FData[-1] := BYTE#16#41;
        FData[0] := BYTE#16#42;
        FData[2] := 120;
        FData[3] := 120;
        FWideData[-1] := WORD#16#0141;
        FWideData[0] := WORD#16#0242;
        FWideData[2] := 120;
        FWideData[3] := 120;
        FEqualExpectedResult := E_Result.Failed;
        FEqualExpectedFinding := TRUE;
        FContainsExpectedResult := E_Result.Passed;
        FContainsExpectedFinding := FALSE;
        FStartsWithExpectedResult := E_Result.Failed;
        FStartsWithExpectedFinding := TRUE;
        FEndsWithExpectedResult := E_Result.Failed;
        FEndsWithExpectedFinding := TRUE;
        FWideEqualExpectedResult := E_Result.Failed;
        FWideEqualExpectedFinding := TRUE;
        FWideContainsExpectedResult := E_Result.Passed;
        FWideContainsExpectedFinding := FALSE;
        FWideStartsWithExpectedResult := E_Result.Failed;
        FWideStartsWithExpectedFinding := TRUE;
        FWideEndsWithExpectedResult := E_Result.Failed;
        FWideEndsWithExpectedFinding := TRUE;
ELSE
    Error(Message := 'Unknown array Assertion scenario.');
    RETURN;
END_CASE;

SelectScenario := TRUE;
END_METHOD

END_FUNCTION_BLOCK

// ---- Framework/Assertions/POU/Arrays/Byte/AssertArrayEqualString_Byte.TcPOU
{region 'Documentation'}
(*!
<summary>Check that the selected array exactly equals the STRING code units.</summary>
<description>

StartIndex is an absolute declared IN index, not an offset. Length selects 1..255
elements; the complete selected range must fit IN. Invalid references or ranges report
Error.

Keep supplied arrays stable for the call. Input data is read, not copied or retained as a
snapshot.

Expected must be nonempty and fit its configured text capacity (otherwise Error). A valid
text longer than the selected array region reports Failed. The array is not zero-terminated or
trimmed; matching is exact and case-sensitive.

The selected array length must equal the text length; trailing padding counts as
data.

</description>
*)
{endregion}
FUNCTION_BLOCK AssertArrayEqualString_Byte EXTENDS AssertionBase
VAR_INPUT
    StartIndex : DINT; //! First selected index in IN; uses the array's declared index range, not a zero-based offset.
    Length : USINT; //! Number of selected array elements, from 1 through 255.
END_VAR
VAR_IN_OUT CONSTANT
    IN : ARRAY[*] OF BYTE; //! Read-only actual data; the selected range must remain stable during the call.
    Expected : STRING(Param_Assertions.AssertionStringLength); //! Nonempty expected text, terminated within the configured capacity; keep stable during the call.
END_VAR

SUPER^();

{region 'Documentation'}
(*!
<summary>Validate references and ranges before exact code-unit comparison.</summary>
*)
{endregion}
METHOD PROTECTED Assert
VAR
    InLowerIndex : DINT;
    InUpperIndex : DINT;
    EndIndex : LINT;
    ExpectedLength : DINT;
    CharacterIndex : DINT;
    InIndex : DINT;
    CandidateOffset : LINT;
    LastCandidateOffset : LINT;
    PatternMatches : BOOL;
    PatternFound : BOOL;
    ExpectedText : STRING(GVL_Constants.AssertionValueLength);
    Message : STRING(GVL_Constants.MessageLength);
END_VAR
VAR CONSTANT
    Terminator : BYTE := 0;
END_VAR
IF NOT EvaluationActive THEN
    RETURN;
END_IF;

IF Result = E_Result.Error THEN
    RETURN;
END_IF;

// C0371: FB inputs are checked before any reference access.
{warning disable C0371}
IF NOT __ISVALIDREF(IN) THEN
    Error(Message := 'Assertion error: IN reference is invalid.');
    RETURN;
END_IF;

IF NOT __ISVALIDREF(Expected) THEN
    Error(Message := 'Assertion error: Expected reference is invalid.');
    RETURN;
END_IF;

IF NOT IsAssertionStringLengthValid(Value := Expected) THEN
    Error(Message := 'Assertion error: Expected exceeds configured STRING length.');
    RETURN;
END_IF;

// SA0175: Exact byte comparison; caller validates termination/capacity and indices stay in bounds.
{analysis -175}
IF Expected[0] = Terminator THEN
{analysis +175}
    Error(Message := 'Assertion error: Expected must not be empty.');
    RETURN;
END_IF;

ExpectedLength := 0;
FOR CharacterIndex := 0 TO UINT_TO_DINT(Param_Assertions.AssertionStringLength) DO
    // SA0175: Exact byte comparison; caller validates termination/capacity and indices stay in bounds.
    {analysis -175}
    IF Expected[CharacterIndex] = Terminator THEN
    {analysis +175}
        ExpectedLength := CharacterIndex;
        EXIT;
    END_IF;
END_FOR;

InLowerIndex := LOWER_BOUND(IN, 1);
InUpperIndex := UPPER_BOUND(IN, 1);
EndIndex := DINT_TO_LINT(StartIndex) + USINT_TO_LINT(Length) - 1;
IF (Length = 0)
    OR (StartIndex < InLowerIndex) OR (StartIndex > InUpperIndex)
    OR (EndIndex > DINT_TO_LINT(InUpperIndex)) THEN
    Message := CONCAT('Assertion error: array range is invalid. StartIndex = ',
        DINT_TO_STRING(StartIndex));
    Message := CONCAT(Message, ', Length = ');
    Message := CONCAT(Message, USINT_TO_STRING(Length));
    Error(Message := Message);
    RETURN;
END_IF;

IF Result = E_Result.Failed THEN
    RETURN;
END_IF;

PatternFound := FALSE;
IF ExpectedLength = USINT_TO_DINT(Length) THEN
    LastCandidateOffset := 0;
    FOR CandidateOffset := 0 TO LastCandidateOffset DO
        PatternMatches := TRUE;
        FOR CharacterIndex := 0 TO ExpectedLength - 1 DO
            InIndex := LINT_TO_DINT(DINT_TO_LINT(StartIndex) + CandidateOffset
                + DINT_TO_LINT(CharacterIndex));
            // SA0175: Exact byte comparison; caller validates termination/capacity and indices stay in bounds.
            {analysis -175}
            IF IN[InIndex] <> Expected[CharacterIndex] THEN
            {analysis +175}
                PatternMatches := FALSE;
                EXIT;
            END_IF;
        END_FOR;
        IF PatternMatches THEN
            PatternFound := TRUE;
            EXIT;
        END_IF;
    END_FOR;
END_IF;

IF NOT PatternFound THEN
    ExpectedText := CreateAssertionTextValue_String(Value := Expected);
    Message := CONCAT('Assertion failed: selected array does not equal Expected = ',
        ExpectedText);
    Message := CONCAT(Message, ', Range = [');
    Message := CONCAT(Message, DINT_TO_STRING(StartIndex));
    Message := CONCAT(Message, '..');
    Message := CONCAT(Message, LINT_TO_STRING(EndIndex));
    Message := CONCAT(Message, '], ExpectedLength = ');
    Message := CONCAT(Message, DINT_TO_STRING(ExpectedLength));
    Message := CONCAT(Message, '.');
    Fail(Message := Message);
    RETURN;
END_IF;

Pass();
{warning restore C0371}
END_METHOD

END_FUNCTION_BLOCK

// ---- Framework/Assertions/POU/Utilities/IsAssertionStringLengthValid.TcPOU
{region 'Documentation'}
(*!
<summary>Checks for a terminator within the configured content capacity, including empty text. Reads at most capacity + 1 code units and stops at the first terminator.</summary>
*)
{endregion}
FUNCTION INTERNAL IsAssertionStringLengthValid : BOOL //! TRUE when a terminator occurs within the configured capacity, including empty text.
VAR_IN_OUT CONSTANT
    Value : STRING(Param_Assertions.AssertionStringLength); //! Read-only text to check for termination within its configured capacity.
END_VAR
VAR
    CharacterIndex : DINT;
END_VAR
VAR CONSTANT
    Terminator : BYTE := 0;
END_VAR

IsAssertionStringLengthValid := FALSE;
FOR CharacterIndex := 0 TO UINT_TO_DINT(Param_Assertions.AssertionStringLength) DO
    // SA0175: Exact byte comparison; caller validates termination/capacity and indices stay in bounds.
    {analysis -175}
    IF Value[CharacterIndex] = Terminator THEN
    {analysis +175}
        IsAssertionStringLengthValid := TRUE;
        RETURN;
    END_IF;
END_FOR;

END_FUNCTION

// ---- Framework/Assertions/POU/Arrays/Byte/AssertArrayContainsString_Byte.TcPOU
{region 'Documentation'}
(*!
<summary>Search the selected array for the contiguous STRING code units.</summary>
<description>

StartIndex is an absolute declared IN index, not an offset. Length selects 1..255
elements; the complete selected range must fit IN. Invalid references or ranges report
Error.

Keep supplied arrays stable for the call. Input data is read, not copied or retained as a
snapshot.

Expected must be nonempty and fit its configured text capacity (otherwise Error). A valid
text longer than the selected array region reports Failed. The array is not zero-terminated or
trimmed; matching is exact and case-sensitive.

</description>
*)
{endregion}
FUNCTION_BLOCK AssertArrayContainsString_Byte EXTENDS AssertionBase
VAR_INPUT
    StartIndex : DINT; //! First selected index in IN; uses the array's declared index range, not a zero-based offset.
    Length : USINT; //! Number of selected array elements, from 1 through 255.
END_VAR
VAR_IN_OUT CONSTANT
    IN : ARRAY[*] OF BYTE; //! Read-only actual data; the selected range must remain stable during the call.
    Expected : STRING(Param_Assertions.AssertionStringLength); //! Nonempty expected text, terminated within the configured capacity; keep stable during the call.
END_VAR

SUPER^();

{region 'Documentation'}
(*!
<summary>Validate references and ranges before exact code-unit comparison.</summary>
*)
{endregion}
METHOD PROTECTED Assert
VAR
    InLowerIndex : DINT;
    InUpperIndex : DINT;
    EndIndex : LINT;
    ExpectedLength : DINT;
    CharacterIndex : DINT;
    InIndex : DINT;
    CandidateOffset : LINT;
    LastCandidateOffset : LINT;
    PatternMatches : BOOL;
    PatternFound : BOOL;
    ExpectedText : STRING(GVL_Constants.AssertionValueLength);
    Message : STRING(GVL_Constants.MessageLength);
END_VAR
VAR CONSTANT
    Terminator : BYTE := 0;
END_VAR
IF NOT EvaluationActive THEN
    RETURN;
END_IF;

IF Result = E_Result.Error THEN
    RETURN;
END_IF;

// C0371: FB inputs are checked before any reference access.
{warning disable C0371}
IF NOT __ISVALIDREF(IN) THEN
    Error(Message := 'Assertion error: IN reference is invalid.');
    RETURN;
END_IF;

IF NOT __ISVALIDREF(Expected) THEN
    Error(Message := 'Assertion error: Expected reference is invalid.');
    RETURN;
END_IF;

IF NOT IsAssertionStringLengthValid(Value := Expected) THEN
    Error(Message := 'Assertion error: Expected exceeds configured STRING length.');
    RETURN;
END_IF;

// SA0175: Exact byte comparison; caller validates termination/capacity and indices stay in bounds.
{analysis -175}
IF Expected[0] = Terminator THEN
{analysis +175}
    Error(Message := 'Assertion error: Expected must not be empty.');
    RETURN;
END_IF;

ExpectedLength := 0;
FOR CharacterIndex := 0 TO UINT_TO_DINT(Param_Assertions.AssertionStringLength) DO
    // SA0175: Exact byte comparison; caller validates termination/capacity and indices stay in bounds.
    {analysis -175}
    IF Expected[CharacterIndex] = Terminator THEN
    {analysis +175}
        ExpectedLength := CharacterIndex;
        EXIT;
    END_IF;
END_FOR;

InLowerIndex := LOWER_BOUND(IN, 1);
InUpperIndex := UPPER_BOUND(IN, 1);
EndIndex := DINT_TO_LINT(StartIndex) + USINT_TO_LINT(Length) - 1;
IF (Length = 0)
    OR (StartIndex < InLowerIndex) OR (StartIndex > InUpperIndex)
    OR (EndIndex > DINT_TO_LINT(InUpperIndex)) THEN
    Message := CONCAT('Assertion error: array range is invalid. StartIndex = ',
        DINT_TO_STRING(StartIndex));
    Message := CONCAT(Message, ', Length = ');
    Message := CONCAT(Message, USINT_TO_STRING(Length));
    Error(Message := Message);
    RETURN;
END_IF;

IF Result = E_Result.Failed THEN
    RETURN;
END_IF;

PatternFound := FALSE;
IF ExpectedLength <= USINT_TO_DINT(Length) THEN
    LastCandidateOffset := USINT_TO_LINT(Length) - DINT_TO_LINT(ExpectedLength);
    FOR CandidateOffset := 0 TO LastCandidateOffset DO
        PatternMatches := TRUE;
        FOR CharacterIndex := 0 TO ExpectedLength - 1 DO
            InIndex := LINT_TO_DINT(DINT_TO_LINT(StartIndex) + CandidateOffset
                + DINT_TO_LINT(CharacterIndex));
            // SA0175: Exact byte comparison; caller validates termination/capacity and indices stay in bounds.
            {analysis -175}
            IF IN[InIndex] <> Expected[CharacterIndex] THEN
            {analysis +175}
                PatternMatches := FALSE;
                EXIT;
            END_IF;
        END_FOR;
        IF PatternMatches THEN
            PatternFound := TRUE;
            EXIT;
        END_IF;
    END_FOR;
END_IF;

IF NOT PatternFound THEN
    ExpectedText := CreateAssertionTextValue_String(Value := Expected);
    Message := CONCAT('Assertion failed: selected array does not contain Expected = ',
        ExpectedText);
    Message := CONCAT(Message, ', Range = [');
    Message := CONCAT(Message, DINT_TO_STRING(StartIndex));
    Message := CONCAT(Message, '..');
    Message := CONCAT(Message, LINT_TO_STRING(EndIndex));
    Message := CONCAT(Message, '], ExpectedLength = ');
    Message := CONCAT(Message, DINT_TO_STRING(ExpectedLength));
    Message := CONCAT(Message, '.');
    Fail(Message := Message);
    RETURN;
END_IF;

Pass();
{warning restore C0371}
END_METHOD

END_FUNCTION_BLOCK

// ---- Framework/Assertions/POU/Arrays/Byte/AssertArrayStartsWithString_Byte.TcPOU
{region 'Documentation'}
(*!
<summary>Check that the selected array starts with the STRING code units.</summary>
<description>

StartIndex is an absolute declared IN index, not an offset. Length selects 1..255
elements; the complete selected range must fit IN. Invalid references or ranges report
Error.

Keep supplied arrays stable for the call. Input data is read, not copied or retained as a
snapshot.

Expected must be nonempty and fit its configured text capacity (otherwise Error). A valid
text longer than the selected array region reports Failed. The array is not zero-terminated or
trimmed; matching is exact and case-sensitive.

</description>
*)
{endregion}
FUNCTION_BLOCK AssertArrayStartsWithString_Byte EXTENDS AssertionBase
VAR_INPUT
    StartIndex : DINT; //! First selected index in IN; uses the array's declared index range, not a zero-based offset.
    Length : USINT; //! Number of selected array elements, from 1 through 255.
END_VAR
VAR_IN_OUT CONSTANT
    IN : ARRAY[*] OF BYTE; //! Read-only actual data; the selected range must remain stable during the call.
    Expected : STRING(Param_Assertions.AssertionStringLength); //! Nonempty expected text, terminated within the configured capacity; keep stable during the call.
END_VAR

SUPER^();

{region 'Documentation'}
(*!
<summary>Validate references and ranges before exact code-unit comparison.</summary>
*)
{endregion}
METHOD PROTECTED Assert
VAR
    InLowerIndex : DINT;
    InUpperIndex : DINT;
    EndIndex : LINT;
    ExpectedLength : DINT;
    CharacterIndex : DINT;
    InIndex : DINT;
    CandidateOffset : LINT;
    LastCandidateOffset : LINT;
    PatternMatches : BOOL;
    PatternFound : BOOL;
    ExpectedText : STRING(GVL_Constants.AssertionValueLength);
    Message : STRING(GVL_Constants.MessageLength);
END_VAR
VAR CONSTANT
    Terminator : BYTE := 0;
END_VAR
IF NOT EvaluationActive THEN
    RETURN;
END_IF;

IF Result = E_Result.Error THEN
    RETURN;
END_IF;

// C0371: FB inputs are checked before any reference access.
{warning disable C0371}
IF NOT __ISVALIDREF(IN) THEN
    Error(Message := 'Assertion error: IN reference is invalid.');
    RETURN;
END_IF;

IF NOT __ISVALIDREF(Expected) THEN
    Error(Message := 'Assertion error: Expected reference is invalid.');
    RETURN;
END_IF;

IF NOT IsAssertionStringLengthValid(Value := Expected) THEN
    Error(Message := 'Assertion error: Expected exceeds configured STRING length.');
    RETURN;
END_IF;

// SA0175: Exact byte comparison; caller validates termination/capacity and indices stay in bounds.
{analysis -175}
IF Expected[0] = Terminator THEN
{analysis +175}
    Error(Message := 'Assertion error: Expected must not be empty.');
    RETURN;
END_IF;

ExpectedLength := 0;
FOR CharacterIndex := 0 TO UINT_TO_DINT(Param_Assertions.AssertionStringLength) DO
    // SA0175: Exact byte comparison; caller validates termination/capacity and indices stay in bounds.
    {analysis -175}
    IF Expected[CharacterIndex] = Terminator THEN
    {analysis +175}
        ExpectedLength := CharacterIndex;
        EXIT;
    END_IF;
END_FOR;

InLowerIndex := LOWER_BOUND(IN, 1);
InUpperIndex := UPPER_BOUND(IN, 1);
EndIndex := DINT_TO_LINT(StartIndex) + USINT_TO_LINT(Length) - 1;
IF (Length = 0)
    OR (StartIndex < InLowerIndex) OR (StartIndex > InUpperIndex)
    OR (EndIndex > DINT_TO_LINT(InUpperIndex)) THEN
    Message := CONCAT('Assertion error: array range is invalid. StartIndex = ',
        DINT_TO_STRING(StartIndex));
    Message := CONCAT(Message, ', Length = ');
    Message := CONCAT(Message, USINT_TO_STRING(Length));
    Error(Message := Message);
    RETURN;
END_IF;

IF Result = E_Result.Failed THEN
    RETURN;
END_IF;

PatternFound := FALSE;
IF ExpectedLength <= USINT_TO_DINT(Length) THEN
    LastCandidateOffset := 0;
    FOR CandidateOffset := 0 TO LastCandidateOffset DO
        PatternMatches := TRUE;
        FOR CharacterIndex := 0 TO ExpectedLength - 1 DO
            InIndex := LINT_TO_DINT(DINT_TO_LINT(StartIndex) + CandidateOffset
                + DINT_TO_LINT(CharacterIndex));
            // SA0175: Exact byte comparison; caller validates termination/capacity and indices stay in bounds.
            {analysis -175}
            IF IN[InIndex] <> Expected[CharacterIndex] THEN
            {analysis +175}
                PatternMatches := FALSE;
                EXIT;
            END_IF;
        END_FOR;
        IF PatternMatches THEN
            PatternFound := TRUE;
            EXIT;
        END_IF;
    END_FOR;
END_IF;

IF NOT PatternFound THEN
    ExpectedText := CreateAssertionTextValue_String(Value := Expected);
    Message := CONCAT('Assertion failed: selected array does not start with Expected = ',
        ExpectedText);
    Message := CONCAT(Message, ', Range = [');
    Message := CONCAT(Message, DINT_TO_STRING(StartIndex));
    Message := CONCAT(Message, '..');
    Message := CONCAT(Message, LINT_TO_STRING(EndIndex));
    Message := CONCAT(Message, '], ExpectedLength = ');
    Message := CONCAT(Message, DINT_TO_STRING(ExpectedLength));
    Message := CONCAT(Message, '.');
    Fail(Message := Message);
    RETURN;
END_IF;

Pass();
{warning restore C0371}
END_METHOD

END_FUNCTION_BLOCK

// ---- Framework/Assertions/POU/Arrays/Byte/AssertArrayEndsWithString_Byte.TcPOU
{region 'Documentation'}
(*!
<summary>Check that the selected array ends with the STRING code units.</summary>
<description>

StartIndex is an absolute declared IN index, not an offset. Length selects 1..255
elements; the complete selected range must fit IN. Invalid references or ranges report
Error.

Keep supplied arrays stable for the call. Input data is read, not copied or retained as a
snapshot.

Expected must be nonempty and fit its configured text capacity (otherwise Error). A valid
text longer than the selected array region reports Failed. The array is not zero-terminated or
trimmed; matching is exact and case-sensitive.

</description>
*)
{endregion}
FUNCTION_BLOCK AssertArrayEndsWithString_Byte EXTENDS AssertionBase
VAR_INPUT
    StartIndex : DINT; //! First selected index in IN; uses the array's declared index range, not a zero-based offset.
    Length : USINT; //! Number of selected array elements, from 1 through 255.
END_VAR
VAR_IN_OUT CONSTANT
    IN : ARRAY[*] OF BYTE; //! Read-only actual data; the selected range must remain stable during the call.
    Expected : STRING(Param_Assertions.AssertionStringLength); //! Nonempty expected text, terminated within the configured capacity; keep stable during the call.
END_VAR

SUPER^();

{region 'Documentation'}
(*!
<summary>Validate references and ranges before exact code-unit comparison.</summary>
*)
{endregion}
METHOD PROTECTED Assert
VAR
    InLowerIndex : DINT;
    InUpperIndex : DINT;
    EndIndex : LINT;
    ExpectedLength : DINT;
    CharacterIndex : DINT;
    InIndex : DINT;
    CandidateOffset : LINT;
    LastCandidateOffset : LINT;
    PatternMatches : BOOL;
    PatternFound : BOOL;
    ExpectedText : STRING(GVL_Constants.AssertionValueLength);
    Message : STRING(GVL_Constants.MessageLength);
END_VAR
VAR CONSTANT
    Terminator : BYTE := 0;
END_VAR
IF NOT EvaluationActive THEN
    RETURN;
END_IF;

IF Result = E_Result.Error THEN
    RETURN;
END_IF;

// C0371: FB inputs are checked before any reference access.
{warning disable C0371}
IF NOT __ISVALIDREF(IN) THEN
    Error(Message := 'Assertion error: IN reference is invalid.');
    RETURN;
END_IF;

IF NOT __ISVALIDREF(Expected) THEN
    Error(Message := 'Assertion error: Expected reference is invalid.');
    RETURN;
END_IF;

IF NOT IsAssertionStringLengthValid(Value := Expected) THEN
    Error(Message := 'Assertion error: Expected exceeds configured STRING length.');
    RETURN;
END_IF;

// SA0175: Exact byte comparison; caller validates termination/capacity and indices stay in bounds.
{analysis -175}
IF Expected[0] = Terminator THEN
{analysis +175}
    Error(Message := 'Assertion error: Expected must not be empty.');
    RETURN;
END_IF;

ExpectedLength := 0;
FOR CharacterIndex := 0 TO UINT_TO_DINT(Param_Assertions.AssertionStringLength) DO
    // SA0175: Exact byte comparison; caller validates termination/capacity and indices stay in bounds.
    {analysis -175}
    IF Expected[CharacterIndex] = Terminator THEN
    {analysis +175}
        ExpectedLength := CharacterIndex;
        EXIT;
    END_IF;
END_FOR;

InLowerIndex := LOWER_BOUND(IN, 1);
InUpperIndex := UPPER_BOUND(IN, 1);
EndIndex := DINT_TO_LINT(StartIndex) + USINT_TO_LINT(Length) - 1;
IF (Length = 0)
    OR (StartIndex < InLowerIndex) OR (StartIndex > InUpperIndex)
    OR (EndIndex > DINT_TO_LINT(InUpperIndex)) THEN
    Message := CONCAT('Assertion error: array range is invalid. StartIndex = ',
        DINT_TO_STRING(StartIndex));
    Message := CONCAT(Message, ', Length = ');
    Message := CONCAT(Message, USINT_TO_STRING(Length));
    Error(Message := Message);
    RETURN;
END_IF;

IF Result = E_Result.Failed THEN
    RETURN;
END_IF;

PatternFound := FALSE;
IF ExpectedLength <= USINT_TO_DINT(Length) THEN
    LastCandidateOffset := USINT_TO_LINT(Length) - DINT_TO_LINT(ExpectedLength);
    FOR CandidateOffset := USINT_TO_LINT(Length) - DINT_TO_LINT(ExpectedLength) TO LastCandidateOffset DO
        PatternMatches := TRUE;
        FOR CharacterIndex := 0 TO ExpectedLength - 1 DO
            InIndex := LINT_TO_DINT(DINT_TO_LINT(StartIndex) + CandidateOffset
                + DINT_TO_LINT(CharacterIndex));
            // SA0175: Exact byte comparison; caller validates termination/capacity and indices stay in bounds.
            {analysis -175}
            IF IN[InIndex] <> Expected[CharacterIndex] THEN
            {analysis +175}
                PatternMatches := FALSE;
                EXIT;
            END_IF;
        END_FOR;
        IF PatternMatches THEN
            PatternFound := TRUE;
            EXIT;
        END_IF;
    END_FOR;
END_IF;

IF NOT PatternFound THEN
    ExpectedText := CreateAssertionTextValue_String(Value := Expected);
    Message := CONCAT('Assertion failed: selected array does not end with Expected = ',
        ExpectedText);
    Message := CONCAT(Message, ', Range = [');
    Message := CONCAT(Message, DINT_TO_STRING(StartIndex));
    Message := CONCAT(Message, '..');
    Message := CONCAT(Message, LINT_TO_STRING(EndIndex));
    Message := CONCAT(Message, '], ExpectedLength = ');
    Message := CONCAT(Message, DINT_TO_STRING(ExpectedLength));
    Message := CONCAT(Message, '.');
    Fail(Message := Message);
    RETURN;
END_IF;

Pass();
{warning restore C0371}
END_METHOD

END_FUNCTION_BLOCK

// ---- Framework/Assertions/POU/Arrays/Word/AssertArrayEqualWString_Word.TcPOU
{region 'Documentation'}
(*!
<summary>Check that the selected array exactly equals the WSTRING code units.</summary>
<description>

StartIndex is an absolute declared IN index, not an offset. Length selects 1..255
elements; the complete selected range must fit IN. Invalid references or ranges report
Error.

Keep supplied arrays stable for the call. Input data is read, not copied or retained as a
snapshot.

Expected must be nonempty and fit its configured text capacity (otherwise Error). A valid
text longer than the selected array region reports Failed. The array is not zero-terminated or
trimmed; matching is exact and case-sensitive.

The selected array length must equal the text length; trailing padding counts as
data.

</description>
*)
{endregion}
FUNCTION_BLOCK AssertArrayEqualWString_Word EXTENDS AssertionBase
VAR_INPUT
    StartIndex : DINT; //! First selected index in IN; uses the array's declared index range, not a zero-based offset.
    Length : USINT; //! Number of selected array elements, from 1 through 255.
END_VAR
VAR_IN_OUT CONSTANT
    IN : ARRAY[*] OF WORD; //! Read-only actual data; the selected range must remain stable during the call.
    Expected : WSTRING(Param_Assertions.AssertionWStringLength); //! Nonempty expected text, terminated within the configured capacity; keep stable during the call.
END_VAR

SUPER^();

{region 'Documentation'}
(*!
<summary>Validate references and ranges before exact code-unit comparison.</summary>
*)
{endregion}
METHOD PROTECTED Assert
VAR
    InLowerIndex : DINT;
    InUpperIndex : DINT;
    EndIndex : LINT;
    ExpectedLength : DINT;
    CharacterIndex : DINT;
    InIndex : DINT;
    CandidateOffset : LINT;
    LastCandidateOffset : LINT;
    PatternMatches : BOOL;
    PatternFound : BOOL;
    ExpectedText : STRING(GVL_Constants.AssertionValueLength);
    Message : STRING(GVL_Constants.MessageLength);
END_VAR
VAR CONSTANT
    Terminator : WORD := 0;
END_VAR
IF NOT EvaluationActive THEN
    RETURN;
END_IF;

IF Result = E_Result.Error THEN
    RETURN;
END_IF;

// C0371: FB inputs are checked before any reference access.
{warning disable C0371}
IF NOT __ISVALIDREF(IN) THEN
    Error(Message := 'Assertion error: IN reference is invalid.');
    RETURN;
END_IF;

IF NOT __ISVALIDREF(Expected) THEN
    Error(Message := 'Assertion error: Expected reference is invalid.');
    RETURN;
END_IF;

IF NOT IsAssertionWStringLengthValid(Value := Expected) THEN
    Error(Message := 'Assertion error: Expected exceeds configured WSTRING length.');
    RETURN;
END_IF;

IF Expected[0] = Terminator THEN
    Error(Message := 'Assertion error: Expected must not be empty.');
    RETURN;
END_IF;

ExpectedLength := 0;
FOR CharacterIndex := 0 TO UINT_TO_DINT(Param_Assertions.AssertionWStringLength) DO
    IF Expected[CharacterIndex] = Terminator THEN
        ExpectedLength := CharacterIndex;
        EXIT;
    END_IF;
END_FOR;

InLowerIndex := LOWER_BOUND(IN, 1);
InUpperIndex := UPPER_BOUND(IN, 1);
EndIndex := DINT_TO_LINT(StartIndex) + USINT_TO_LINT(Length) - 1;
IF (Length = 0)
    OR (StartIndex < InLowerIndex) OR (StartIndex > InUpperIndex)
    OR (EndIndex > DINT_TO_LINT(InUpperIndex)) THEN
    Message := CONCAT('Assertion error: array range is invalid. StartIndex = ',
        DINT_TO_STRING(StartIndex));
    Message := CONCAT(Message, ', Length = ');
    Message := CONCAT(Message, USINT_TO_STRING(Length));
    Error(Message := Message);
    RETURN;
END_IF;

IF Result = E_Result.Failed THEN
    RETURN;
END_IF;

